// TIA Portal project "batch Steam cooker V2" (V19)

(* hardware
DEVICE "S7-1200 station_1"  S7-1200 Station
   slot 0: "Rack_0"  S7-1200 Rack  Rack  V1.0
   slot 1: "PLC_1"  CPU 1214C AC/DC/Rly  6ES7 214-1BG40-0XB0  V4.5
DEVICE "HMI_2"  TP700 Comfort
   slot 0: "HMI_2"  TP700 Comfort  6AV2 124-0GC01-0AX0  17.0.0.0
   slot 1: "HMI_RT_2"  TP700 Comfort  6AV2 124-0GC01-0AX0  17.0.0.0
   slot 5: "HMI_2.IE_CP_1"  PROFINET Interface  17.0.0.0
      slot 1: "PROFINET Interface_1"  PROFINET Interface
         slot 1: "Port_1"  Port
         slot 2: "Port_2"  Port
   slot 7: "HMI_2.MPI/DP_CP_1"  MPI/DP Interface  17.0.0.0
*)

// ===== PLC "PLC_1"  CPU 1214C AC/DC/Rly =====

VAR_GLOBAL   // PLC tag table "Default tag table"
   "Vacuum Pump Starter" AT %Q4.0 : Bool;
   "Steam Regulator" AT %Q4.1 : Bool;
   "Cooling Water Valve" AT %Q4.2 : Bool;
   "Green Light" AT %Q3.0 : Bool;
   "Red Light" AT %Q3.2 : Bool;
   "Yellow Light" AT %Q3.1 : Bool;
   "Alarm_Word" AT %MW3 : Int;
   "Tag_1" AT %M3.0 : Bool;
   "Tag_2" AT %M3.1 : Bool;
   "Tag_3" AT %M3.6 : Bool;
   "Tag_4" AT %M3.7 : Bool;
   "Tag_5" AT %M4.0 : Bool;
   "Tag_6" AT %M4.1 : Bool;
   "Tag_7" AT %M3.2 : Bool;
   "Tag_8" AT %M3.3 : Bool;
   "Tag_9" AT %M3.4 : Bool;
   "Tag_10" AT %M3.5 : Bool;
   "Acknowledge_Word" AT %MW4 : Int;
   "Acknowledge bit" AT %M5.0 : Bool;
END_VAR

VAR_GLOBAL   // PLC tag table "IO_Inputs"
   "Door Lock FB" AT %I0.1 : Bool;
   "Manhole Closed FB" AT %I0.2 : Bool;
   "Manhole Open FB" AT %I0.3 : Bool;
   "Water Level FB" AT %I0.4 : Bool;
   "Door Interlock" AT %I0.5 : Bool;
   "Emergency Stop" AT %I0.7 : Bool;
   "Pressure Input" AT %ID68 : Real;
   "Temperature Input" AT %ID64 : Real;
   "Water Flow Input" AT %ID72 : Real;
END_VAR

VAR_GLOBAL   // PLC tag table "IO_Outputs"
   "V1 Output" AT %Q0.0 : Bool;
   "V2 Output" AT %Q0.1 : Bool;
   "V3 Output" AT %Q0.2 : Bool;
   "V9" AT %Q1.0 : Bool;
   "V8" AT %Q0.7 : Bool;
   "V7" AT %Q0.6 : Bool;
   "V6" AT %Q0.5 : Bool;
   "V5" AT %Q0.4 : Bool;
   "V4" AT %Q0.3 : Bool;
   "Motor Run Output" AT %Q2.0 : Bool;
   "Motor Direction Output" AT %Q2.1 : Bool;
END_VAR

VAR_GLOBAL CONSTANT   // PLC tag table "Const"
   "cIdle" : Int := 50;
   "cLock" : Int := 15;
   "cAddWater" : Int := 1;
   "cOpenMH" : Int := 2;
   "cWaitMat" : Int := 3;
   "cCloseMH" : Int := 4;
   "cColdMix" : Int := 5;
   "cHeat" : Int := 6;
   "cCook" : Int := 7;
   "cConfDis" : Int := 10;
   "cDisch" : Int := 11;
   "cFinal" : Int := 12;
END_VAR

TYPE "UDT_Recipe_Production"
   STRUCT
      Recipe_Name : String := 'DEFAULT';   // Recipe identification name
      Recipe_Number : UInt := 1;   // Recipe ID number (1-99)
      Heating_Temp_Phase1 : Real := 80.0;   // Cooking temperature setpoint (°C)
      Adding_Water1_QTY : Real := 100.0;   // First water addition quantity (Liters)
      Cold_Mix_Time : Time := T#300S;   // Cold mix time before heating (seconds)
      Cooking_Time_Phase1 : Time := T#1800S;   // Cooking time after temp reached (seconds)
      Compensation_Time : Time := T#600S;   // Additional processing time (seconds)
      Discharge_Time : Time;   // Auto discharge time (0=manual only)
      Water_Flow_Timeout : Time := T#120S;   // Water addition timeout
      Manhole_Open_Time : Time :=  T#30S;   // Manhole opening timeout
      Manhole_Close_Time : Time :=  T#30S;   // Manhole closing timeout
      Steam_Ramp_Rate : Real := 5.0;   // Steam valve opening rate %/sec
      Vacuum_Enable : Bool := true;   // Enable vacuum during cooking
      Final_Temp_Target : Real := 75.0;   // Final product temperature (°C)
      Product_Type : UInt := 1;   // Product type (1=Soft, 2=Hard, 3=Special)
      Batch_Size_kg : Real := 300.0;
   END_STRUCT;
END_TYPE

TYPE "UDT_Motor_Command"
   STRUCT
      Priority : UInt := 0;   // Command priority (1=Auto, 2=Func, 3=Man)
      Start_Man : Bool;
      Start_Func : Bool;
      Start_Auto : Bool;
      Stop : Bool;
      Reset : Bool;
      Pulse_Enable : Bool;
      Discharge_Mode : Bool;
      Enable : Bool;
      Direction : Int;
      Speed_SP_pct : Real;   // Speed setpoint %
   END_STRUCT;
END_TYPE

TYPE "UDT_Motor_Config"
   STRUCT
      Motor_Name : String;
      Max_Speed_pct : Real := 100.0;
      Min_Speed_pct : Real := 0.0;
      Start_Timeout : Time := T#10S;
      Stop_Timeout : Time := T#5S ;
      Rev_Dwell : Time := T#2S ;   // Direction change dwell
      T_Fwd : Time := T#30S ;
      T_Hold : Time := T#5S ;
      T_Bwd : Time := T#20S ;
      Disch_Speed_pct : Real := 25.0;
      Acceleration_Time : Time := T#3S;
      Deceleration_Time : Time := T#3S;
      Interlock_Used : Bool := TRUE;
      Motor_Type : UInt := 1;
      Rated_Speed_RPM : Real;
      Rated_Power_kW : Real;
   END_STRUCT;
END_TYPE

TYPE "UDT_Motor_Status"
   STRUCT
      Running : Bool;   // Motor is running
      Fault : Bool;
      Fault_Code : UInt;
      Direction : UInt;   // Direction (0=Stop, 1=Fwd, 2=Rev)
      State : UInt;   // State (0=Stop, 1=Fwd, 2=Hold, 3=Bwd)
      Source : UInt;   // Command source (0=None, 1=Auto, 2=Func, 3=Man)
      Ready : Bool;
      Position_pct : Real;   // Position feedback %
      Speed_Actual_pct : Real;
      Runtime_Hours : Real;
      Start_Count : UDInt;
      R_Fwd : Bool;
      R_Rev : Bool;
      RDwell_Q : Bool;
   END_STRUCT;
END_TYPE

TYPE "UDT_Motor_Outputs"
   STRUCT
      Q_Run : Bool;
      Q_DirFwd : Bool;
      Q_Stop : Bool;
      Contactor_Main : Bool;
      Contactor_Star : Bool;
      Contactor_Delta : Bool;
      Brake_Release : Bool;
      Alarm_Output : Bool;
      Status_LED : UInt;
      AO_SpeedPct : Real;
      AO_Torque : Real;
   END_STRUCT;
END_TYPE

TYPE "UDT_Motor_Interlocks"
   STRUCT
      Permissive : Bool := true;   // General permissive
      OOS : Bool;   // Out of service
      E_Stop : Bool;
      Drive_Ready : Bool;   // Drive ready feedback
      Drive_Fault : Bool;
      Temperature_OK : Bool := true;
      Vibration_OK : Bool := true;
      Overcurrent_OK : Bool := true;
      Door_Closed : Bool := TRUE;
      Guard_OK : Bool := TRUE;
      Lubrication_OK : Bool := TRUE;
      Cooling_OK : Bool := TRUE;
      Local_Stop : Bool;
      Drive_Running : Bool;
      Overload : Bool;
      VFD_Fault : Bool;
   END_STRUCT;
END_TYPE

TYPE "UDT_Motor"
   STRUCT
      Command : "UDT_Motor_Command";
      Outputs : "UDT_Motor_Outputs";   // Physical outputs
      Config : "UDT_Motor_Config";
      Status : "UDT_Motor_Status";
      Interlocks : "UDT_Motor_Interlocks";
   END_STRUCT;
END_TYPE

TYPE "UDT_Valve_Command"
   STRUCT
      Priority : UInt;
      Open_Man : Bool;
      Open_Auto : Bool;
      Close_Auto : Bool;
      Close_Man : Bool;
      Open_Func : Bool;
      Close_Func : Bool;
      Reset : Bool;
      Emergency_Close : Bool;
   END_STRUCT;
END_TYPE

TYPE "UDT_Valve_Config"
   STRUCT
      Valve_Type : UInt := 1;
      Valve_Name : String;
      Travel_Timeout : Time := T#30ms;
      Stroke_Time : Time := T#15ms;
      Position_Tolerance : Real := 2.0;
      Min_Position : Real;
      Max_Position : Real := 100.0;
      Fail_Position : UInt;
      TwoCoils : Bool;
      Actuator_Type : UInt := 1;
      Feedback_Type : UInt := 1;
      Service_Hours : Real;
      Interlock_Used : Bool := True;
      Fail_Safe_Position : Bool;
      Open_Time : Time;
      Close_Time : Time;
   END_STRUCT;
END_TYPE

TYPE "UDT_Valve_Status"
   STRUCT
      Fault : Bool;
      Fault_Code : UInt;
      State : UInt;   // State (0=Stop, 1=Fwd, 2=Hold, 3=Bwd)
      Source : UInt;   // Command source (0=None, 1=Auto, 2=Func, 3=Man)
      Ready : Bool;
      Moving : Bool;
      At_Position : Bool;
      Travel_Time : Time;
      Operation_Count : UDInt;
      Position_Actual_pct : Real;   // Position feedback %
      Runtime_Hours : Real;
      Limit_Open : Bool;
      Limit_Closed : Bool;
      Open : Bool;
      Closed : Bool;
   END_STRUCT;
END_TYPE

TYPE "UDT_Valve_Outputs"
   STRUCT
      Q_Run : Bool;
      Q_Open : Bool;
      Q_Close : Bool;
      Solenoid_A : Bool;
      Solenoid_B : Bool;
      Motor_CW : Bool;
      Motor_CCW : Bool;
      Brake_Release : Bool;
      Status_LED : Bool;
      Alarm_Output : Bool;
      AO_Position_pct : Real;
   END_STRUCT;
END_TYPE

TYPE "UDT_Valve_Interlocks"
   STRUCT
      Permissive : Bool := true;   // General permissive
      OOS : Bool;   // Out of service
      E_Stop : Bool;
      Process_Temp_OK : Bool := true;
      Local_Isolation : Bool;
      Process_Pressure_OK : Bool := TRUE        ;
      Upstream_OK : Bool := TRUE        ;
      Downstream_OK : Bool := TRUE        ;
      Interlock_Chain : Bool := TRUE        ;
      Maintenance_Lock : Bool;
      Air_Pressure_OK : Bool := TRUE        ;
      Power_Available : Bool := TRUE        ;
   END_STRUCT;
END_TYPE

TYPE "UDT_Valve"
   STRUCT
      Command : "UDT_Valve_Command";
      Config : "UDT_Valve_Config";
      Status : "UDT_Valve_Status";
      Outputs : "UDT_Valve_Outputs";
      Interlocks : "UDT_Valve_Interlocks";
      Open_Auto : Bool;
      Priority : UInt;
      Reset : Bool;
      Open_Man : Bool;
      Close_Man : Bool;
      Open_Func : Bool;
      Close_Func : Bool;
      Close_Auto : Bool;
      Position_SP_pct : Real;
      Enable : Bool;
      Emergency_Close : Bool;
   END_STRUCT;
END_TYPE

TYPE "UDT_Recipe_Screw"
   STRUCT
      Forward_Speed_pct : Real := 75.0;   // Forward screw speed %
      Backward_Speed_pct : Real := 50.0;
      Reverse_Speed_pct : Real := 50.0;
      Forward_Run_Time : Time := T#30S ;   // Forward running time (pulsing)
      Backward_Run_Time : Time := T#20S ;
      Hold_Time : Time := T#10S ;   // Hold time between direction changes
      Pause_Time : Time := T#5S ;   // Pause between pulse cycles
      Direction_Change_Delay : Time := T#2S;   // Delay between direction changes
      Screw_Ramp_Time : Time := T#3S;   // Speed ramp up/down time
      Max_Runtime_Continuous : Time := T#600S;   // Max continuous runtime before pause
      Discharge_Speed_pct : Real := 25.0;   // Screw speed during discharge %
      Cold_Mix_Speed_pct : Real := 60.0;   // Speed during cold mixing %
      Cook_Mix_Speed_pct : Real := 80.0;   // Speed during cooking phase %
      Pulse_Enable_ColdMix : Bool := TRUE;   // Enable pulsing during cold mix
      Pulse_Enable_Cooking : Bool := TRUE;
      Pulse_Enable_Discharge : Bool;
      Pulse_Time_On : Time;
      Pulse_Time_Off : Time;
   END_STRUCT;
END_TYPE

TYPE "UDT_Recipe_Temperature"
   STRUCT
      Heat_Setpoint_Phase1 : Real := 80.0;
      Heat_Setpoint_Phase2 : Real := 85.0;
      Heat_Deadband : Real := 2.0;
      Heat_Rate_Limit : Real := 2.0;
      Cool_Setpoint : Real := 60.0;
      Cool_Rate_Limit : Real := 1.0;
      Steam_Pressure_Max : Real := 6.0;
      Steam_Pressure_Min : Real := 2.0;
      Temp_Alarm_High : Real := 95.0;
      Temp_Alarm_Low : Real := 40.0;
      Temp_Sensor_Timeout : Time := T#10S;
      Heat_Timeout : Time := T#1800S;
      Cool_Timeout : Time := T#900S;
      Overtemp_Shutdown : Real := 100.0;
      Cool_Deadband : Real;
   END_STRUCT;
END_TYPE

TYPE "UDT_Recipe_Vacuum"
   STRUCT
      Vacuum_Setpoint_mbar : Real := 500.0;   // Vacuum setpoint (mbar absolute)
      Vacuum_Tolerance : Real := 50.0;   // Vacuum tolerance (±mbar)
      Vacuum_Offset_pct : Real := 5.0;   // Hysteresis offset percentage
      Pump_Start_Delay : Time := T#5S;   // Pump start delay after valve open
      Pump_Stop_Delay : Time := T#10S;   // Pump stop delay after valve close
      Max_Vacuum_Time : Time := T#3600S;   // aximum continuous vacuum time
      Vacuum_Break_Pressure : Real := 900.0;   // Vacuum break pressure (mbar)
      Leak_Test_Time : Time := T#60S;   // Vacuum leak test duration
      Leak_Test_Tolerance : Real := 10.0;   // Acceptable leak rate (mbar/min)
      Emergency_Break_Enable : Bool := TRUE;   // Enable emergency vacuum break
      Cooling_Vacuum_Enable : Bool := TRUE;   // Enable vacuum during cooling
      Cooking_Vacuum_Enable : Bool;
      Vacuum_Pump_Timeout : Time := T#30S;   // Vacuum pump start timeout
      Pressure_Sensor_Timeout : Time := T#10S;   // Pressure sensor timeout
      Min_Vacuum_Quality : Real := 100.0;   // Minimum vacuum level (mbar)
   END_STRUCT;
END_TYPE

TYPE "UDT_Recipe_Complete"
   STRUCT
      Production : "UDT_Recipe_Production";   // Production parameters
      Screw : "UDT_Recipe_Screw";
      Temperature : "UDT_Recipe_Temperature";
      Vacuum : "UDT_Recipe_Vacuum";
      Recipe_Valid : Bool;
      Recipe_Locked : Bool;
      Creation_Date : DTL;
      Modified_Date : DTL;
      Created_By : String := 'SYSTEM';
      Modified_By : String := 'SYSTEM';
      Recipe_Version : Real := 1.0;
      Recipe_Notes : String;
   END_STRUCT;
END_TYPE

TYPE "UDT_Process_Status"
   STRUCT
      Current_Step : UInt := 50;
      Step_Name : String := 'IDLE';
      Phase_Name : String := 'IDLE';
      Phase_Active : UInt;   // Active phase (0=Idle, 1=Prep, 2=Mix, 3=Cook, 4=Discharge)
      Current_Phase : UInt;
      Time_Remaining : Time;
      Time_Elapsed : Time;
      Total_Batch_Time : Time;
      Step_Progress_pct : Real;
      Batch_Progress_pct : Real;
      Temp_Actual : Real := 25.0;
      Temp_Setpoint : Real;
      Pressure_Actual : Real := 1013.0;
      Pressure_Setpoint : Real;   // Current pressure setpoint (mbar)
      Water_Level_Actual : Real;
      Water_Level_Target : Real;
      Screw_Speed_Actual : Real;
      Screw_Speed_Setpoint : Real;   // Screw speed setpoint %
      Batch_Number : UInt := 1;   // Current water level (L)
      Recipe_Active : UInt := 1;
      Process_Running : Bool;
      Process_Paused : Bool;
      Process_Complete : Bool;
      Process_Aborted : Bool;
      Fault_Active : Bool;   // System fault active flag
      Emergency_Stop : Bool;   // Emergency stop active flag
      Operator_Present : Bool;   // Operator attention required
      System_Ready : Bool;
      Overall_Progress : Real;
      Individual_Discharge_Active : Bool;
   END_STRUCT;
END_TYPE

TYPE "UDT_Process_HMI"
   STRUCT
      Start_Production : Bool;
      Stop_Production : Bool;
      Reset_System : Bool;
      Reset_p_s : Bool;
      Abort_Process : Bool;
      Acknowledge_Alarms : Bool;
      RawMaterial_OK : Bool;
      Manhole_Secured_OK : Bool;
      Discharge_Ready_OK : Bool;
      Quality_Check_OK : Bool;
      Cleaning_Complete_OK : Bool;
      Recipe_Selected : UInt := 1;
      Load_Recipe : Bool;
      Save_Recipe : Bool;
      Recipe_Edit_Mode : Bool;
      Recipe_Backup : Bool;
      Recipe_Restore : Bool;
      Manual_ON : Array[0..15] of Bool;   // Manual ON commands [V1-V9, R1, Aux1-5]
      Manual_OFF : Array[0..15] of Bool;
      Auto_Mode : Array[0..15] of Bool;
      Temp_Override_Enable : Bool;
      Temp_Override_Value : Real;
      Speed_Override_Enable : Bool;
      Speed_Override_Value : Real;
      Time_Override_Enable : Bool;
      Time_Override_Factor : Real := 1.0;
      Operator_ID : String := 'UNKNOWN';
      Shift_ID : UInt := 1;
      Production_Mode : UInt := 1;   // Mode (1=Auto, 2=Manual, 3=Test)
      System_Ready : Bool;
      Maintenance_Mode : Bool;
      Individual_Discharge_Button : Bool;
   END_STRUCT;
END_TYPE

TYPE "UDT_Process_IO"
   STRUCT
      FS_Water_Flow : Bool;
      LS1_Discharge_Locked : Bool;
      LS2_Manhole_Closed : Bool;
      LS3_Manhole_Opened : Bool;
      LL_Water_Level : Bool;
      ES_Emergency_Stop : Bool;
      PS_Steam_Pressure_OK : Bool;
      PS_Air_Pressure_OK : Bool;
      TS_Steam_Temperature_OK : Bool;
      Door_Interlock_OK : Bool;
      Guard_Switch_OK : Bool;
      Door_Locked_FB : Bool;
      Door_Unlocked_FB : Bool;
      Water_Level_FB : Bool;
      Manhole_Open_FB : Bool;
      Manhole_Closed_FB : Bool;
      AI_Temperature : Real := 25.0;
      AI_Pressure : Real := 1013.0;
      AI_Steam_Pressure : Real;
      AI_Water_Flow : Real;
      AI_Steam_Flow : Real;
      AI_Vacuum_Level : Real := 1013.0;
      AI_Motor_Current : Real;
      AI_Motor_Power : Real;
      DO_Alarm_Horn : Bool;
      DO_Status_Green : Bool;
      DO_Status_Yellow : Bool;
      DO_Status_Red : Bool;
      DO_Vacuum_Pump : Bool;   // Vacuum pump starter (K1)
      DO_Steam_Regulator_En : Bool;
      DO_Cooling_Water : Bool;
      DO_Process_Light : Bool;
      AO_Steam_Regulator : Real;
      AO_Cooling_Control : Real;
      AO_Process_Speed : Real;
   END_STRUCT;
END_TYPE

DATA_BLOCK "DB_Recipes"   // DB1
{ S7_Optimized_Access := 'TRUE' }
VERSION : 0.1
   VAR
      Recipes : Array[1..10] of "UDT_Recipe_Complete";   // Recipe storage array (1-10)
      Active_Recipe : "UDT_Recipe_Complete";   // Currently loaded recipe
      Default_Recipe : "UDT_Recipe_Complete";   // Factory default recipe
   END_VAR
BEGIN
   Default_Recipe.Production.Recipe_Name := 'DEFAULT_CHEESE';
   Default_Recipe.Production.Batch_Size_kg := 1000.0;
   Default_Recipe.Production.Adding_Water1_QTY := 100.0;
   Default_Recipe.Production.Water_Flow_Timeout := T#120S;
   Default_Recipe.Production.Cold_Mix_Time := T#300S;
   Default_Recipe.Production.Cooking_Time_Phase1 := T#1800S;
   Default_Recipe.Production.Heating_Temp_Phase1 := 80.0;
   Default_Recipe.Screw.Cold_Mix_Speed_pct := 60.0;
   Default_Recipe.Screw.Cook_Mix_Speed_pct := 80.0;
   Default_Recipe.Screw.Discharge_Speed_pct := 25.0;
   Default_Recipe.Temperature.Heat_Setpoint_Phase1 := 80.0;
   Default_Recipe.Temperature.Heat_Deadband := 2.0;
   Default_Recipe.Temperature.Heat_Timeout := T#1800S;
   Default_Recipe.Recipe_Valid := TRUE;
   Default_Recipe.Production.Recipe_Number := 1;
   Default_Recipe.Production.Manhole_Open_Time := T#30S;
   Default_Recipe.Production.Manhole_Close_Time := T#30S;
   Default_Recipe.Screw.Pulse_Enable_ColdMix := TRUE;
   Default_Recipe.Screw.Pulse_Enable_Cooking := TRUE;
   Default_Recipe.Vacuum.Vacuum_Setpoint_mbar := 500.0;
   Default_Recipe.Vacuum.Vacuum_Tolerance := 50.0;
   Default_Recipe.Vacuum.Cooking_Vacuum_Enable := FALSE;
   Active_Recipe.Production.Water_Flow_Timeout := T#10S;
   Active_Recipe.Production.Compensation_Time := T#6S;
   Active_Recipe.Production.Cooking_Time_Phase1 := T#10S;
   Active_Recipe.Production.Cold_Mix_Time := T#20S;
   Active_Recipe.Production.Discharge_Time := T#6ms;
   Active_Recipe.Vacuum.Cooking_Vacuum_Enable := TRUE;
END_DATA_BLOCK

DATA_BLOCK "FB_Process_Main_DB"   // DB2
{ S7_Optimized_Access := 'TRUE' }
VERSION : 0.1
// stored: InstanceOfName FB_Process_Main
"FB_Process_Main"
BEGIN
END_DATA_BLOCK

DATA_BLOCK "FB_Motor_VFD_DB_1"   // DB3
{ S7_Optimized_Access := 'TRUE' }
VERSION : 0.1
// stored: InstanceOfName FB_Motor_VFD
"FB_Motor_VFD"
BEGIN
END_DATA_BLOCK

DATA_BLOCK "FB_Motor_VFD_DB"   // DB13
{ S7_Optimized_Access := 'TRUE' }
VERSION : 0.1
// stored: InstanceOfName FB_Motor_VFD
"FB_Motor_VFD"
BEGIN
END_DATA_BLOCK

DATA_BLOCK "ALarms"   // DB14
{ S7_Optimized_Access := 'TRUE' }
VERSION : 0.1
   VAR
      Alarms : UInt;
   END_VAR
BEGIN
END_DATA_BLOCK

DATA_BLOCK "FB_Valve_DO_DB"   // DB15
{ S7_Optimized_Access := 'TRUE' }
VERSION : 0.1
// stored: InstanceOfName FB_Valve_DO
"FB_Valve_DO"
BEGIN
END_DATA_BLOCK

DATA_BLOCK "DB_Motors"   // DB18
{ S7_Optimized_Access := 'TRUE' }
VERSION : 0.1
   VAR RETAIN
      Motors : Array[1..1] of "UDT_Motor";   // Motor control array - =Screw Motor
   END_VAR
BEGIN
   Motors[1].Config.Motor_Name := 'SCREW_MOTOR';
   Motors[1].Config.Max_Speed_pct := 1800.0;
   Motors[1].Config.Rated_Speed_RPM := 1800.0;
   Motors[1].Config.Rated_Power_kW := 15.0;
   Motors[1].Config.Acceleration_Time := T#10S;
   Motors[1].Config.Rev_Dwell := T#2S;
   Motors[1].Config.Disch_Speed_pct := 25.0;
   Motors[1].Config.Start_Timeout := T#10S;
   Motors[1].Config.T_Fwd := T#30S;
   Motors[1].Config.T_Hold := T#5S;
   Motors[1].Config.T_Bwd := T#20S;
END_DATA_BLOCK

DATA_BLOCK "DB_Valves"   // DB19
{ S7_Optimized_Access := 'TRUE' }
VERSION : 0.1
   VAR
      Valves : Array[1..9] of "UDT_Valve";   // Valve control array - =V1 Manhole, =V2 CIP, ..., =V9 Vacuum Cooling
   END_VAR
BEGIN
   Valves[1].Config.Valve_Name := 'V1_MANHOLE';
   Valves[2].Config.Valve_Name := 'V2_CIP';
   Valves[3].Config.Valve_Name := 'V3_DISCHARGE_UNLOCK';
   Valves[4].Config.Valve_Name := 'V4_DISCHARGE';
   Valves[5].Config.Valve_Name := 'V5_WATER';
   Valves[6].Config.Valve_Name := 'V6_STEAM';
   Valves[7].Config.Valve_Name := 'V7_EVACUATION';
   Valves[8].Config.Valve_Name := 'V8_VACUUM';
   Valves[9].Config.Valve_Name := 'V9_VACUUM_COOLING';
   Valves[1].Config.Travel_Timeout := T#30S;
   Valves[2].Config.Travel_Timeout := T#15S;
   Valves[3].Config.Travel_Timeout := T#30S;
   Valves[4].Config.Travel_Timeout := T#20S;
   Valves[5].Config.Travel_Timeout := T#15S;
   Valves[6].Config.Travel_Timeout := T#10S;
   Valves[7].Config.Travel_Timeout := T#15S;
   Valves[8].Config.Travel_Timeout := T#20S;
   Valves[9].Config.Travel_Timeout := T#15S;
END_DATA_BLOCK

DATA_BLOCK "DB_Test_Motors"   // DB20
{ S7_Optimized_Access := 'FALSE' }
VERSION : 0.1
   VAR
      ff : Int;
   END_VAR
BEGIN
END_DATA_BLOCK

DATA_BLOCK "DB_Process"   // DB21
{ S7_Optimized_Access := 'FALSE' }
VERSION : 0.1
   VAR
      Status : "UDT_Process_Status";   // current process
      HMI : "UDT_Process_HMI";
      IO : "UDT_Process_IO";
      Timers : Array[1..10] of TON_TIME;
      Counters : Array[1..5] of CTU_INT;
   END_VAR
BEGIN
   Status.Current_Step := 50;
   Status.Step_Name := 'IDLE';
   Status.Batch_Number := 1;
   Status.Recipe_Active := 1;
   HMI.Shift_ID := 1;
   HMI.Operator_ID := 'OPERATOR';
   IO.AI_Pressure := 1000.0;
   IO.AI_Steam_Pressure := 25.0;
   IO.Manhole_Open_FB := true;
END_DATA_BLOCK

FUNCTION_BLOCK "FB_Valve_DO"   // FB1, LAD
{ S7_Optimized_Access := 'TRUE' }
VERSION : 0.1
   VAR_INPUT
      AutoCmd : Bool;   // from automatic sequence (open=TRUE)
      FuncCmd : Bool;   // from Function screens
      ManCmd : Bool;   // from Manual page (your ON/OFF button drives this)
      OOS : Bool;   // Out Of Service; forces closed
      Permissive : Bool;   // E‑Stop OK, interlocks OK
      FbOpen : Bool;   // optional open limit switch
      FbClosed : Bool;   // optional closed limit switch
      TwoCoils : Bool;   // TRUE = separate open/close coils; FALSE = single coil
      T_Stroke : Time := T#3S;   // normal movement time (e.g., T#5S)
      T_Timeout : Time := T#6S;   // fault timeout (e.g., T#10S)
   END_VAR
   VAR_OUTPUT
      Q_Open : Bool;   // open (or single) coil
      Q_Close : Bool;   // close coil (only used if TwoCoils=TRUE)
      Ready : Bool;
      FaultTO : Bool;
      FaultFB : Bool;
      Source : UInt;   // 1 Auto, 2 Func, 3 Man
      Status : UInt;   // 0 Unknown, 1 Closed, 2 Opening, 3 Open, 4 Closing, 5 Fault
   END_VAR
   VAR
      Cmd_DesiredOpen_raw : Bool;
      Cmd_DesiredOpen_OK : Bool;
      Req_Open : Bool;
      Req_Close : Bool;
      St_Opening : Bool;
      St_Closing : Bool;
      St_Open : Bool;
      St_Closed : Bool;
      St_Moving : Bool;
      Open_Reached : Bool;
      Close_Reached : Bool;
      FaultLatched : Bool;
      TON_Move : TON_TIME;
      TON_Timeout : TON_TIME;
   END_VAR
   VAR_TEMP
      MoveEnable : Bool;
   END_VAR
BEGIN

REGION Network 1: Conflict for feedback
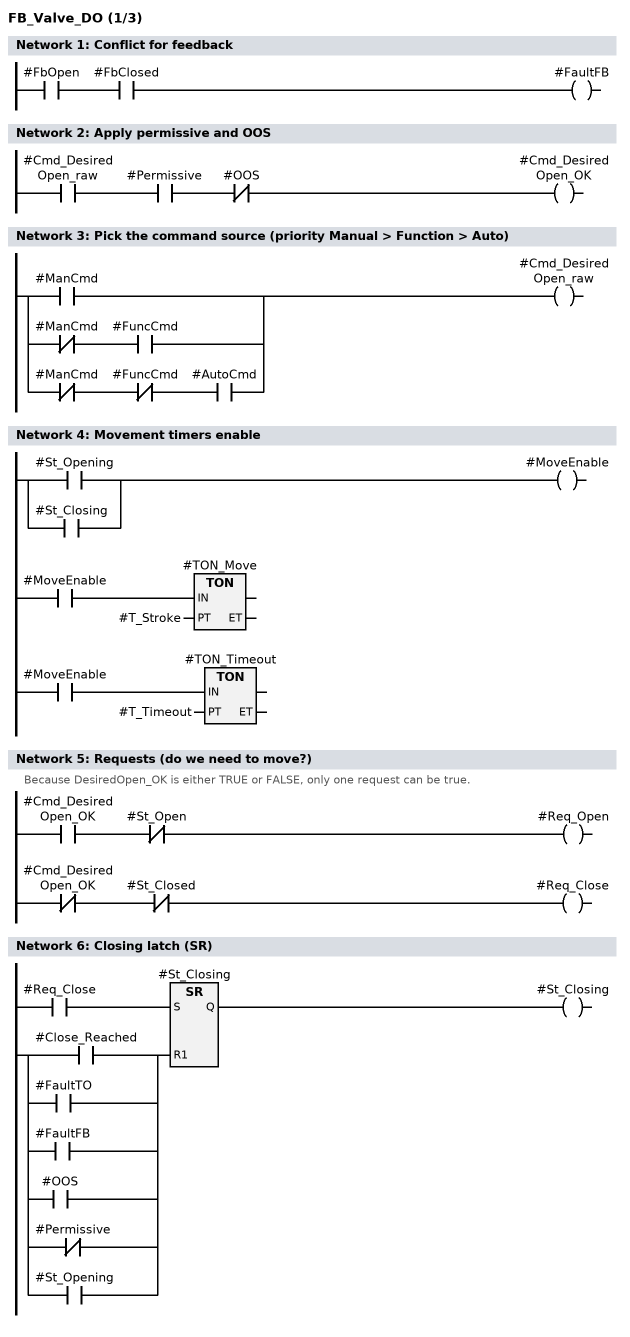
   RUNG wire#powerrail
      Contact( #FbOpen )
      Contact( #FbClosed )
      Coil( #FaultFB )
   END_RUNG
   // the same network as SCL:
   #FaultFB := #FbOpen AND #FbClosed;
END_REGION

REGION Network 2: Apply permissive and OOS
   RUNG wire#powerrail
      Contact( #Cmd_DesiredOpen_raw )
      Contact( #Permissive )
      I_Contact( #OOS )
      Coil( #Cmd_DesiredOpen_OK )
   END_RUNG
   // the same network as SCL:
   #Cmd_DesiredOpen_OK := #Cmd_DesiredOpen_raw AND #Permissive AND NOT #OOS;
END_REGION

REGION Network 3: Pick the command source (priority Manual > Function > Auto)
   RUNG wire#powerrail
      Contact( #ManCmd )
      wire#w1
      Coil( #Cmd_DesiredOpen_raw )
   END_RUNG
   RUNG wire#powerrail
      I_Contact( #ManCmd )
      Contact( #FuncCmd )
   END_RUNG wire#w1
   RUNG wire#powerrail
      I_Contact( #ManCmd )
      I_Contact( #FuncCmd )
      Contact( #AutoCmd )
   END_RUNG wire#w1
   // the same network as SCL:
   #Cmd_DesiredOpen_raw := #ManCmd OR (NOT #ManCmd AND #FuncCmd) OR (NOT #ManCmd AND NOT #FuncCmd AND #AutoCmd);
END_REGION

REGION Network 4: Movement timers enable
   #MoveEnable := #St_Opening OR #St_Closing;
   #TON_Move(IN := #MoveEnable, PT := #T_Stroke);   // TON
   #TON_Timeout(IN := #MoveEnable, PT := #T_Timeout);   // TON
END_REGION

REGION Network 5: Requests (do we need to move?)
   // Because DesiredOpen_OK is either TRUE or FALSE, only one request can be true.
   RUNG wire#powerrail
      Contact( #Cmd_DesiredOpen_OK )
      I_Contact( #St_Open )
      Coil( #Req_Open )
   END_RUNG
   RUNG wire#powerrail
      I_Contact( #Cmd_DesiredOpen_OK )
      I_Contact( #St_Closed )
      Coil( #Req_Close )
   END_RUNG
   // the same network as SCL:
   #Req_Open := #Cmd_DesiredOpen_OK AND NOT #St_Open;
   #Req_Close := NOT #Cmd_DesiredOpen_OK AND NOT #St_Closed;
END_REGION

REGION Network 6: Closing latch (SR)
   RUNG wire#powerrail
      Contact( #Req_Close )
      S_SR(operand := #St_Closing, r1 := wire#w1)
      Coil( #St_Closing )
   END_RUNG
   RUNG wire#powerrail
      Contact( #Close_Reached )
   END_RUNG wire#w1
   RUNG wire#powerrail
      Contact( #FaultTO )
   END_RUNG wire#w1
   RUNG wire#powerrail
      Contact( #FaultFB )
   END_RUNG wire#w1
   RUNG wire#powerrail
      Contact( #OOS )
   END_RUNG wire#w1
   RUNG wire#powerrail
      I_Contact( #Permissive )
   END_RUNG wire#w1
   RUNG wire#powerrail
      Contact( #St_Opening )
   END_RUNG wire#w1
   // the same network as SCL:
   IF #Req_Close THEN
       #St_Closing := TRUE;   // SR flip-flop
   END_IF;
   IF #Close_Reached OR #FaultTO OR #FaultFB OR #OOS OR NOT #Permissive OR #St_Opening THEN
       #St_Closing := FALSE;
   END_IF;
   #St_Closing := #St_Closing;
END_REGION

REGION Network 7: Latch “Opening” (SR)
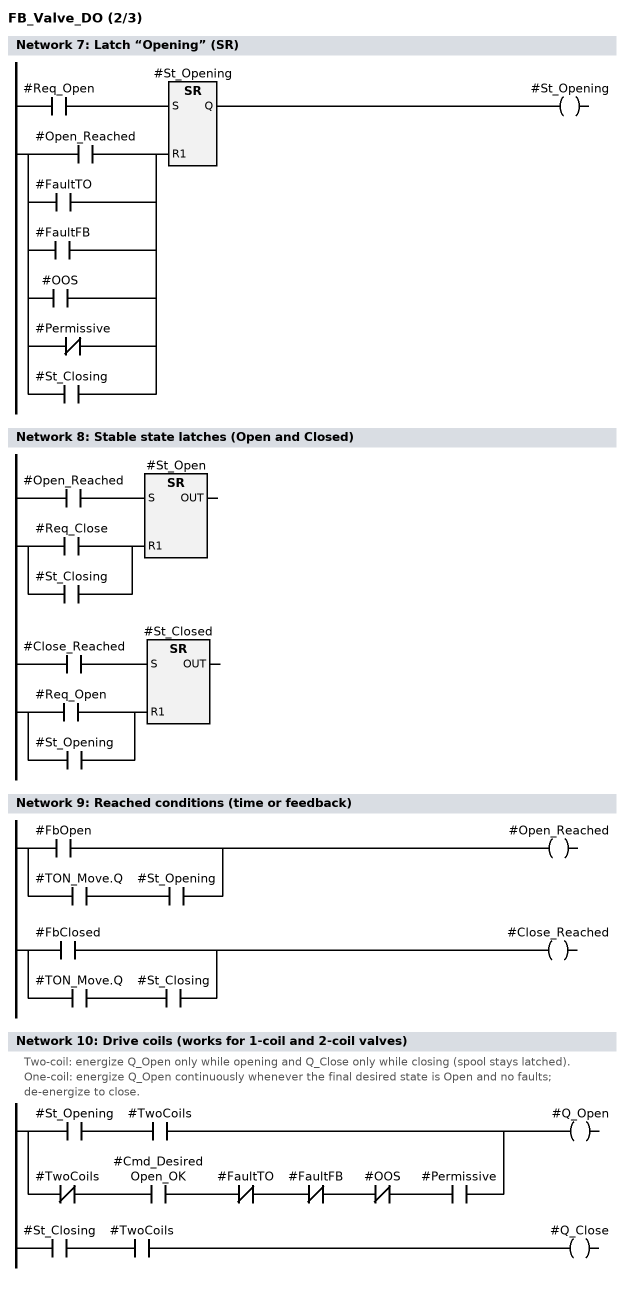
   RUNG wire#powerrail
      Contact( #Req_Open )
      S_SR(operand := #St_Opening, r1 := wire#w1)
      Coil( #St_Opening )
   END_RUNG
   RUNG wire#powerrail
      Contact( #Open_Reached )
   END_RUNG wire#w1
   RUNG wire#powerrail
      Contact( #FaultTO )
   END_RUNG wire#w1
   RUNG wire#powerrail
      Contact( #FaultFB )
   END_RUNG wire#w1
   RUNG wire#powerrail
      Contact( #OOS )
   END_RUNG wire#w1
   RUNG wire#powerrail
      I_Contact( #Permissive )
   END_RUNG wire#w1
   RUNG wire#powerrail
      Contact( #St_Closing )
   END_RUNG wire#w1
   // the same network as SCL:
   IF #Req_Open THEN
       #St_Opening := TRUE;   // SR flip-flop
   END_IF;
   IF #Open_Reached OR #FaultTO OR #FaultFB OR #OOS OR NOT #Permissive OR #St_Closing THEN
       #St_Opening := FALSE;
   END_IF;
   #St_Opening := #St_Opening;
END_REGION

REGION Network 8: Stable state latches (Open and Closed)
   RUNG wire#powerrail
      Contact( #Open_Reached )
      S_SR(operand := #St_Open, r1 := wire#w1)
   END_RUNG
   RUNG wire#powerrail
      Contact( #Req_Close )
   END_RUNG wire#w1
   RUNG wire#powerrail
      Contact( #St_Closing )
   END_RUNG wire#w1
   RUNG wire#powerrail
      Contact( #Close_Reached )
      S_SR(operand := #St_Closed, r1 := wire#w2)
   END_RUNG
   RUNG wire#powerrail
      Contact( #Req_Open )
   END_RUNG wire#w2
   RUNG wire#powerrail
      Contact( #St_Opening )
   END_RUNG wire#w2
   // the same network as SCL:
   IF #Open_Reached THEN
       #St_Open := TRUE;   // SR flip-flop
   END_IF;
   IF #Req_Close OR #St_Closing THEN #St_Open := FALSE; END_IF;
   IF #Close_Reached THEN
       #St_Closed := TRUE;   // SR flip-flop
   END_IF;
   IF #Req_Open OR #St_Opening THEN #St_Closed := FALSE; END_IF;
END_REGION

REGION Network 9: Reached conditions (time or feedback)
   RUNG wire#powerrail
      Contact( #FbOpen )
      wire#w1
      Coil( #Open_Reached )
   END_RUNG
   RUNG wire#powerrail
      Contact( #TON_Move.Q )
      Contact( #St_Opening )
   END_RUNG wire#w1
   RUNG wire#powerrail
      Contact( #FbClosed )
      wire#w2
      Coil( #Close_Reached )
   END_RUNG
   RUNG wire#powerrail
      Contact( #TON_Move.Q )
      Contact( #St_Closing )
   END_RUNG wire#w2
   // the same network as SCL:
   #Open_Reached := #FbOpen OR (#TON_Move.Q AND #St_Opening);
   #Close_Reached := #FbClosed OR (#TON_Move.Q AND #St_Closing);
END_REGION

REGION Network 10: Drive coils (works for 1‑coil and 2‑coil valves)
   // Two‑coil: energize Q_Open only while opening and Q_Close only while closing (spool stays latched).
   // One‑coil: energize Q_Open continuously whenever the final desired state is Open and no faults; de‑energize to close.
   RUNG wire#powerrail
      Contact( #St_Opening )
      Contact( #TwoCoils )
      wire#w1
      Coil( #Q_Open )
   END_RUNG
   RUNG wire#powerrail
      I_Contact( #TwoCoils )
      Contact( #Cmd_DesiredOpen_OK )
      I_Contact( #FaultTO )
      I_Contact( #FaultFB )
      I_Contact( #OOS )
      Contact( #Permissive )
   END_RUNG wire#w1
   RUNG wire#powerrail
      Contact( #St_Closing )
      Contact( #TwoCoils )
      Coil( #Q_Close )
   END_RUNG
   // the same network as SCL:
   #Q_Open := (#St_Opening AND #TwoCoils) OR (NOT #TwoCoils AND #Cmd_DesiredOpen_OK AND NOT #FaultTO AND NOT #FaultFB AND NOT #OOS AND #Permissive);
   #Q_Close := #St_Closing AND #TwoCoils;
END_REGION

REGION Network 11: Ready flag
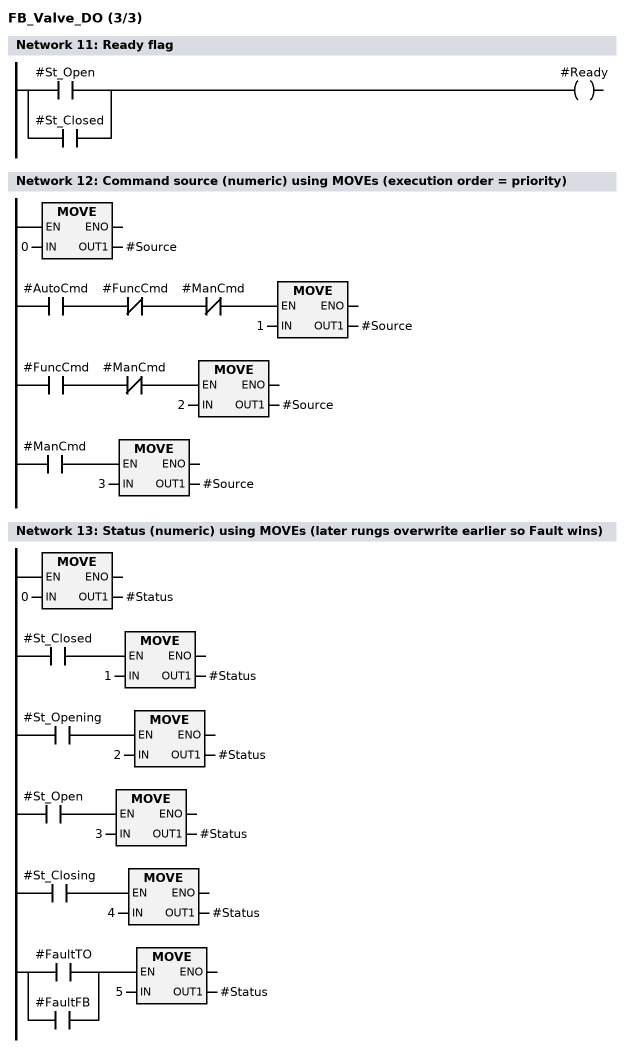
   RUNG wire#powerrail
      Contact( #St_Open )
      wire#w1
      Coil( #Ready )
   END_RUNG
   RUNG wire#powerrail
      Contact( #St_Closed )
   END_RUNG wire#w1
   // the same network as SCL:
   #Ready := #St_Open OR #St_Closed;
END_REGION

REGION Network 12: Command source (numeric) using MOVEs (execution order = priority)
   RUNG wire#powerrail
      Move(in := 0, out1 => #Source)
   END_RUNG
   RUNG wire#powerrail
      Contact( #AutoCmd )
      I_Contact( #FuncCmd )
      I_Contact( #ManCmd )
      Move(in := 1, out1 => #Source)
   END_RUNG
   RUNG wire#powerrail
      Contact( #FuncCmd )
      I_Contact( #ManCmd )
      Move(in := 2, out1 => #Source)
   END_RUNG
   RUNG wire#powerrail
      Contact( #ManCmd )
      Move(in := 3, out1 => #Source)
   END_RUNG
   // the same network as SCL:
   #Source := 0;
   IF #AutoCmd AND NOT #FuncCmd AND NOT #ManCmd THEN #Source := 1; END_IF;
   IF #FuncCmd AND NOT #ManCmd THEN #Source := 2; END_IF;
   IF #ManCmd THEN #Source := 3; END_IF;
END_REGION

REGION Network 13: Status (numeric) using MOVEs (later rungs overwrite earlier so Fault wins)
   RUNG wire#powerrail
      Move(in := 0, out1 => #Status)
   END_RUNG
   RUNG wire#powerrail
      Contact( #St_Closed )
      Move(in := 1, out1 => #Status)
   END_RUNG
   RUNG wire#powerrail
      Contact( #St_Opening )
      Move(in := 2, out1 => #Status)
   END_RUNG
   RUNG wire#powerrail
      Contact( #St_Open )
      Move(in := 3, out1 => #Status)
   END_RUNG
   RUNG wire#powerrail
      Contact( #St_Closing )
      Move(in := 4, out1 => #Status)
   END_RUNG
   RUNG wire#powerrail
      Contact( #FaultTO )
      wire#w1
      Move(in := 5, out1 => #Status)
   END_RUNG
   RUNG wire#powerrail
      Contact( #FaultFB )
   END_RUNG wire#w1
   // the same network as SCL:
   #Status := 0;
   IF #St_Closed THEN #Status := 1; END_IF;
   IF #St_Opening THEN #Status := 2; END_IF;
   IF #St_Open THEN #Status := 3; END_IF;
   IF #St_Closing THEN #Status := 4; END_IF;
   IF #FaultTO OR #FaultFB THEN #Status := 5; END_IF;
END_REGION
END_FUNCTION_BLOCK

FUNCTION_BLOCK "FB_Motor_VFD"   // FB2, LAD
{ S7_Optimized_Access := 'TRUE' }
VERSION : 0.1
   VAR_INPUT
      Start_Auto : Bool;
      Start_Func : Bool;
      Start_Man : Bool;
      OOS : Bool;
      RevDwell : Time := T#2S;
      Permissive : Bool := true;
      PulseEnable : Bool;   // TRUE = do Fwd/Hold/Bwd pulsing
      T_Fwd : Time := T#8S;
      T_Hold : Time := T#2S;
      T_Bwd : Time := T#6S;
      DischargeMode : Bool;   // TRUE = forward only
      SpeedSP_pct : Real;   // 0..100, normal speed
      DischSpeed_pct : Real;   // 0..100, used when DischargeMode=TRUE
      DriveReady : Bool;   // optional, from VFD
      DriveFault : Bool;   // optional, from VFD
      StartTimeout : Time := T#5S;
   END_VAR
   VAR_OUTPUT
      Q_Run : Bool;   // to RUN relay or PN run bit
      Q_DirFwd : Bool;   // TRUE = forward, FALSE = reverse
      AO_SpeedPct : Real;   // speed command 0..100%
      Running : Bool;
      Direction : UInt;   // 0 Stop, 1 Fwd, 2 Bwd
      Fault : Bool;
      FaultCode : UInt;   // 0 ok, 1 timeout, 2 drive fault, 3 permissive/OOS
      Source : UInt;   // 1 Auto, 2 Func, 3 Man
      R_Fwd : Bool;
      R_Rev : Bool;
      State : UInt;   // 0 Stop, 1 Fwd, 2 Hold, 3 Bwd (for HMI)
      RDwell_Q : Bool;
   END_VAR
   VAR
      Start_Prio : Bool;
      RunCmd : Bool;
      Start_OK : Bool;
      RStart : R_TRIG;
      St_Fwd : Bool;
      St_Hold : Bool;
      St_Bwd : Bool;
      Tmr_Fwd : TON_TIME;
      Tmr_Hold : TON_TIME;
      Tmr_Bwd : TON_TIME;
      Tmr_Dwell : TON_TIME;
      DwellActive : Bool;
      PrevDirFwd : Bool;
      Tmr_Start : TON_TIME;
      StartRise : Bool;
      PulseActive : Bool;
      RDwell : R_TRIG;
      FDwell : F_TRIG;
      ChangePulse : Bool;
      DwellRun : Bool;
      Start_Raw : Bool;
      DirFwdCmd : Bool;
   END_VAR
BEGIN

REGION Network 1: Command priority (Man > Func > Auto) → Start_Raw
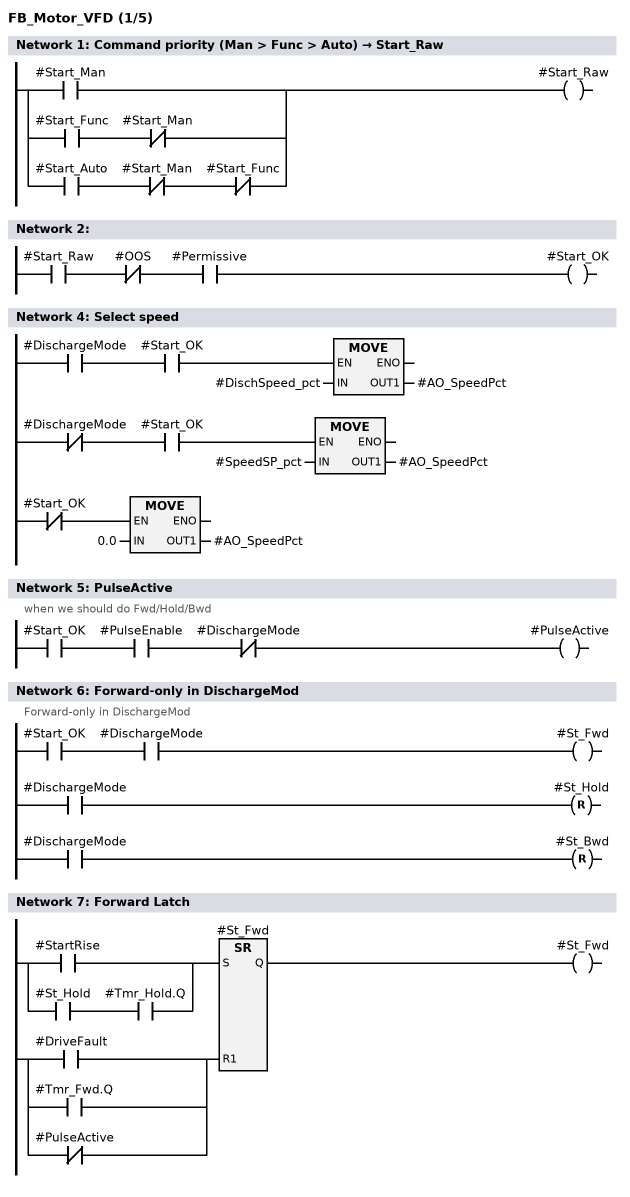
   RUNG wire#powerrail
      Contact( #Start_Man )
      wire#w1
      Coil( #Start_Raw )
   END_RUNG
   RUNG wire#powerrail
      Contact( #Start_Func )
      I_Contact( #Start_Man )
   END_RUNG wire#w1
   RUNG wire#powerrail
      Contact( #Start_Auto )
      I_Contact( #Start_Man )
      I_Contact( #Start_Func )
   END_RUNG wire#w1
   // the same network as SCL:
   #Start_Raw := #Start_Man OR (#Start_Func AND NOT #Start_Man) OR (#Start_Auto AND NOT #Start_Man AND NOT #Start_Func);
END_REGION

REGION Network 2
   RUNG wire#powerrail
      Contact( #Start_Raw )
      I_Contact( #OOS )
      Contact( #Permissive )
      Coil( #Start_OK )
   END_RUNG
   // the same network as SCL:
   #Start_OK := #Start_Raw AND NOT #OOS AND #Permissive;
END_REGION

REGION Network 3 (SCL)
   // CORRECT:
   #RStart(CLK := #Start_OK);
   #StartRise := #RStart.Q;
END_REGION

REGION Network 4: Select speed
   RUNG wire#powerrail
      Contact( #DischargeMode )
      Contact( #Start_OK )
      Move(in := #DischSpeed_pct, out1 => #AO_SpeedPct)
   END_RUNG
   RUNG wire#powerrail
      I_Contact( #DischargeMode )
      Contact( #Start_OK )
      Move(in := #SpeedSP_pct, out1 => #AO_SpeedPct)
   END_RUNG
   RUNG wire#powerrail
      I_Contact( #Start_OK )
      Move(in := 0.0, out1 => #AO_SpeedPct)
   END_RUNG
   // the same network as SCL:
   IF #DischargeMode AND #Start_OK THEN #AO_SpeedPct := #DischSpeed_pct; END_IF;
   IF NOT #DischargeMode AND #Start_OK THEN #AO_SpeedPct := #SpeedSP_pct; END_IF;
   IF NOT #Start_OK THEN #AO_SpeedPct := 0.0; END_IF;
END_REGION

REGION Network 5: PulseActive
   // when we should do Fwd/Hold/Bwd
   RUNG wire#powerrail
      Contact( #Start_OK )
      Contact( #PulseEnable )
      I_Contact( #DischargeMode )
      Coil( #PulseActive )
   END_RUNG
   // the same network as SCL:
   #PulseActive := #Start_OK AND #PulseEnable AND NOT #DischargeMode;
END_REGION

REGION Network 6: Forward-only in DischargeMod
   // Forward-only in DischargeMod
   RUNG wire#powerrail
      Contact( #Start_OK )
      Contact( #DischargeMode )
      Coil( #St_Fwd )
   END_RUNG
   RUNG wire#powerrail
      Contact( #DischargeMode )
      R_Coil( #St_Hold )
   END_RUNG
   RUNG wire#powerrail
      Contact( #DischargeMode )
      R_Coil( #St_Bwd )
   END_RUNG
   // the same network as SCL:
   #St_Fwd := #Start_OK AND #DischargeMode;
   IF #DischargeMode THEN
       #St_Hold := FALSE;
       #St_Bwd := FALSE;
   END_IF;
END_REGION

REGION Network 7: Forward Latch
   RUNG wire#powerrail
      Contact( #StartRise )
      wire#w1
      S_SR(operand := #St_Fwd, r1 := wire#w2)
      Coil( #St_Fwd )
   END_RUNG
   RUNG wire#powerrail
      Contact( #St_Hold )
      Contact( #Tmr_Hold.Q )
   END_RUNG wire#w1
   RUNG wire#powerrail
      Contact( #DriveFault )
   END_RUNG wire#w2
   RUNG wire#powerrail
      Contact( #Tmr_Fwd.Q )
   END_RUNG wire#w2
   RUNG wire#powerrail
      I_Contact( #PulseActive )
   END_RUNG wire#w2
   // the same network as SCL:
   IF #StartRise OR (#St_Hold AND #Tmr_Hold.Q) THEN
       #St_Fwd := TRUE;   // SR flip-flop
   END_IF;
   IF #DriveFault OR #Tmr_Fwd.Q OR NOT #PulseActive THEN #St_Fwd := FALSE; END_IF;
   #St_Fwd := #St_Fwd;
END_REGION

REGION Network 8: Hold Latch
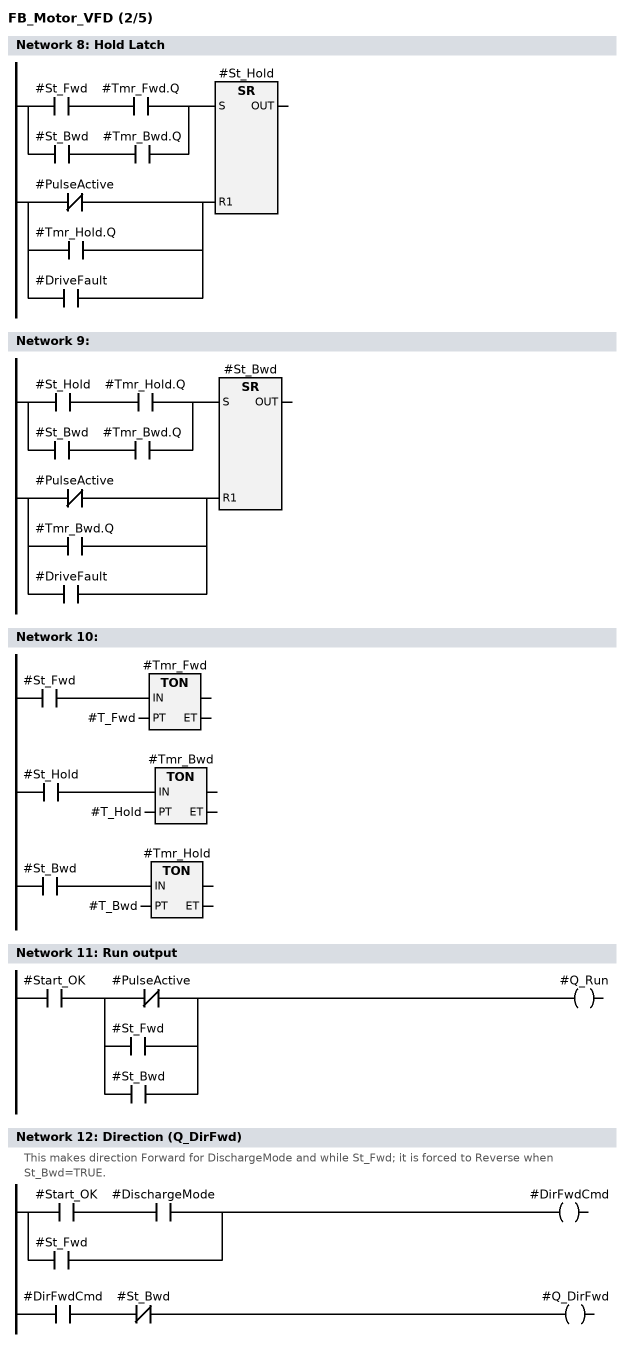
   RUNG wire#powerrail
      Contact( #St_Fwd )
      Contact( #Tmr_Fwd.Q )
      wire#w1
      S_SR(operand := #St_Hold, r1 := wire#w2)
   END_RUNG
   RUNG wire#powerrail
      Contact( #St_Bwd )
      Contact( #Tmr_Bwd.Q )
   END_RUNG wire#w1
   RUNG wire#powerrail
      I_Contact( #PulseActive )
   END_RUNG wire#w2
   RUNG wire#powerrail
      Contact( #Tmr_Hold.Q )
   END_RUNG wire#w2
   RUNG wire#powerrail
      Contact( #DriveFault )
   END_RUNG wire#w2
   // the same network as SCL:
   IF (#St_Fwd AND #Tmr_Fwd.Q) OR (#St_Bwd AND #Tmr_Bwd.Q) THEN
       #St_Hold := TRUE;   // SR flip-flop
   END_IF;
   IF NOT #PulseActive OR #Tmr_Hold.Q OR #DriveFault THEN #St_Hold := FALSE; END_IF;
END_REGION

REGION Network 9
   RUNG wire#powerrail
      Contact( #St_Hold )
      Contact( #Tmr_Hold.Q )
      wire#w1
      S_SR(operand := #St_Bwd, r1 := wire#w2)
   END_RUNG
   RUNG wire#powerrail
      Contact( #St_Bwd )
      Contact( #Tmr_Bwd.Q )
   END_RUNG wire#w1
   RUNG wire#powerrail
      I_Contact( #PulseActive )
   END_RUNG wire#w2
   RUNG wire#powerrail
      Contact( #Tmr_Bwd.Q )
   END_RUNG wire#w2
   RUNG wire#powerrail
      Contact( #DriveFault )
   END_RUNG wire#w2
   // the same network as SCL:
   IF (#St_Hold AND #Tmr_Hold.Q) OR (#St_Bwd AND #Tmr_Bwd.Q) THEN
       #St_Bwd := TRUE;   // SR flip-flop
   END_IF;
   IF NOT #PulseActive OR #Tmr_Bwd.Q OR #DriveFault THEN #St_Bwd := FALSE; END_IF;
END_REGION

REGION Network 10
   #Tmr_Fwd(IN := #St_Fwd, PT := #T_Fwd);   // TON
   #Tmr_Bwd(IN := #St_Hold, PT := #T_Hold);   // TON
   #Tmr_Hold(IN := #St_Bwd, PT := #T_Bwd);   // TON
END_REGION

REGION Network 11: Run output
   RUNG wire#powerrail
      Contact( #Start_OK )
      wire#w1
      I_Contact( #PulseActive )
      wire#w2
      Coil( #Q_Run )
   END_RUNG
   RUNG wire#w1
      Contact( #St_Fwd )
   END_RUNG wire#w2
   RUNG wire#w1
      Contact( #St_Bwd )
   END_RUNG wire#w2
   // the same network as SCL:
   #Q_Run := #Start_OK AND (NOT #PulseActive OR #St_Fwd OR #St_Bwd);
END_REGION

REGION Network 12: Direction (Q_DirFwd)
   // This makes direction Forward for DischargeMode and while St_Fwd; it is forced to Reverse when St_Bwd=TRUE.
   RUNG wire#powerrail
      Contact( #Start_OK )
      Contact( #DischargeMode )
      wire#w1
      Coil( #DirFwdCmd )
   END_RUNG
   RUNG wire#powerrail
      Contact( #St_Fwd )
   END_RUNG wire#w1
   RUNG wire#powerrail
      Contact( #DirFwdCmd )
      I_Contact( #St_Bwd )
      Coil( #Q_DirFwd )
   END_RUNG
   // the same network as SCL:
   #DirFwdCmd := (#Start_OK AND #DischargeMode) OR #St_Fwd;
   #Q_DirFwd := #DirFwdCmd AND NOT #St_Bwd;
END_REGION

REGION Network 13: Detect change of direction
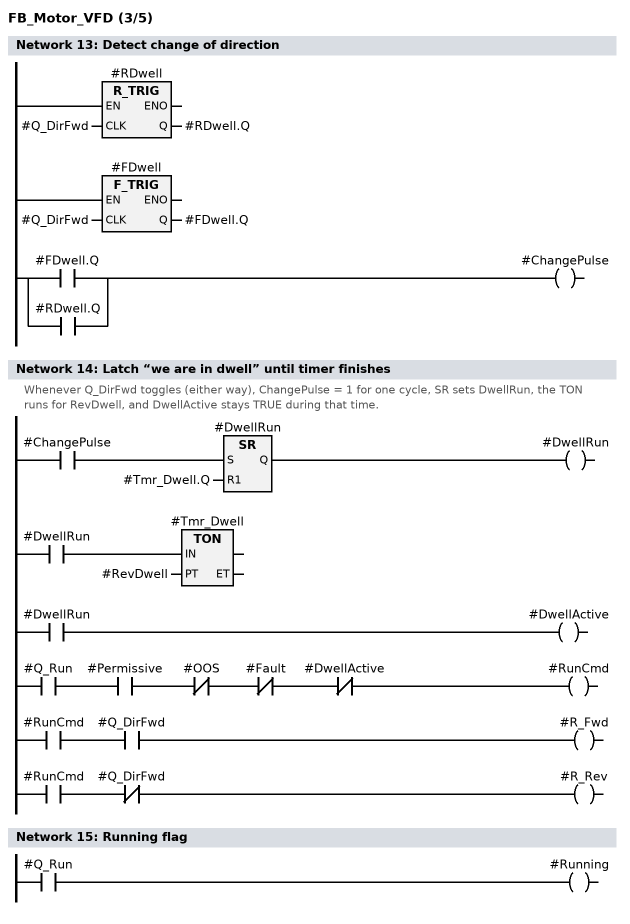
   #RDwell(CLK := #Q_DirFwd, Q => #RDwell.Q);   // R_TRIG
   #FDwell(CLK := #Q_DirFwd, Q => #FDwell.Q);   // F_TRIG
   #ChangePulse := #FDwell.Q OR #RDwell.Q;
END_REGION

REGION Network 14: Latch “we are in dwell” until timer finishes
   // Whenever Q_DirFwd toggles (either way), ChangePulse = 1 for one cycle, SR sets DwellRun, the TON runs for RevDwell, and DwellActive stays TRUE during that time.
   IF #ChangePulse THEN
       #DwellRun := TRUE;   // SR flip-flop
   END_IF;
   IF #Tmr_Dwell.Q THEN #DwellRun := FALSE; END_IF;
   #DwellRun := #DwellRun;
   #Tmr_Dwell(IN := #DwellRun, PT := #RevDwell);   // TON
   #DwellActive := #DwellRun;
   #RunCmd := #Q_Run AND #Permissive AND NOT #OOS AND NOT #Fault AND NOT #DwellActive;
   #R_Fwd := #RunCmd AND #Q_DirFwd;
   #R_Rev := #RunCmd AND NOT #Q_DirFwd;
END_REGION

REGION Network 15: Running flag
   RUNG wire#powerrail
      Contact( #Q_Run )
      Coil( #Running )
   END_RUNG
   // the same network as SCL:
   #Running := #Q_Run;
END_REGION

REGION Network 16: Start timeout and Drive faults
   // if you don’t have DriveReady wiring yet, set DriveReady=TRUE when you CALL the FB so the start timeout won’t trigger.
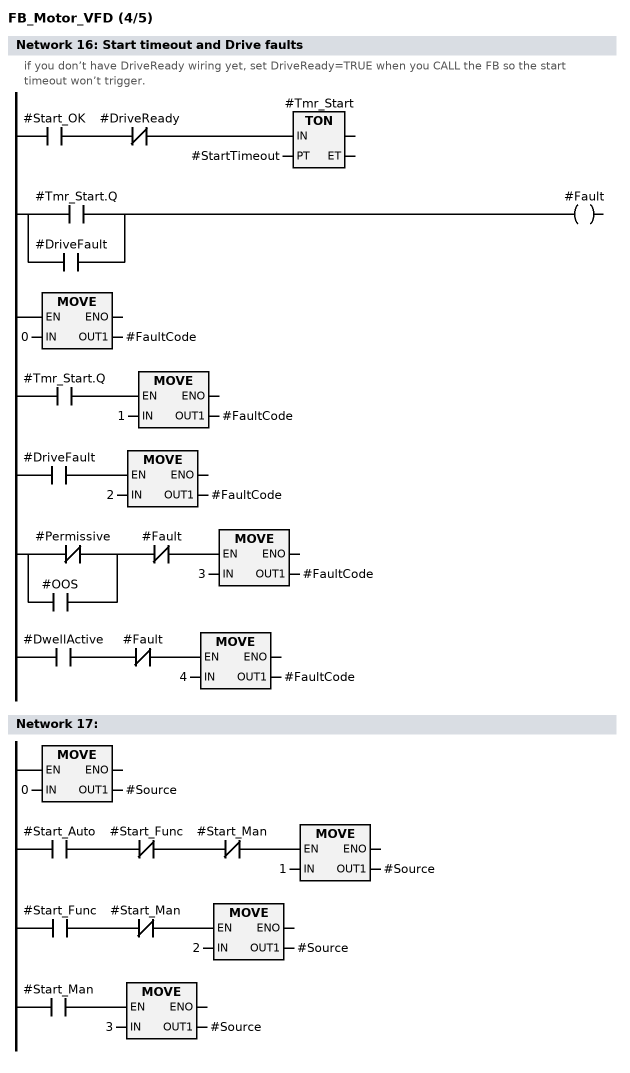
   #Tmr_Start(IN := #Start_OK AND NOT #DriveReady, PT := #StartTimeout);   // TON
   #Fault := #Tmr_Start.Q OR #DriveFault;
   #FaultCode := 0;
   IF #Tmr_Start.Q THEN #FaultCode := 1; END_IF;
   IF #DriveFault THEN #FaultCode := 2; END_IF;
   IF (NOT #Permissive OR #OOS) AND NOT #Fault THEN #FaultCode := 3; END_IF;
   IF #DwellActive AND NOT #Fault THEN #FaultCode := 4; END_IF;
END_REGION

REGION Network 17
   RUNG wire#powerrail
      Move(in := 0, out1 => #Source)
   END_RUNG
   RUNG wire#powerrail
      Contact( #Start_Auto )
      I_Contact( #Start_Func )
      I_Contact( #Start_Man )
      Move(in := 1, out1 => #Source)
   END_RUNG
   RUNG wire#powerrail
      Contact( #Start_Func )
      I_Contact( #Start_Man )
      Move(in := 2, out1 => #Source)
   END_RUNG
   RUNG wire#powerrail
      Contact( #Start_Man )
      Move(in := 3, out1 => #Source)
   END_RUNG
   // the same network as SCL:
   #Source := 0;
   IF #Start_Auto AND NOT #Start_Func AND NOT #Start_Man THEN #Source := 1; END_IF;
   IF #Start_Func AND NOT #Start_Man THEN #Source := 2; END_IF;
   IF #Start_Man THEN #Source := 3; END_IF;
END_REGION

REGION Network 18: State
   // for HMI: 0 Stop, 1 Fwd, 2 Hold, 3 Bwd
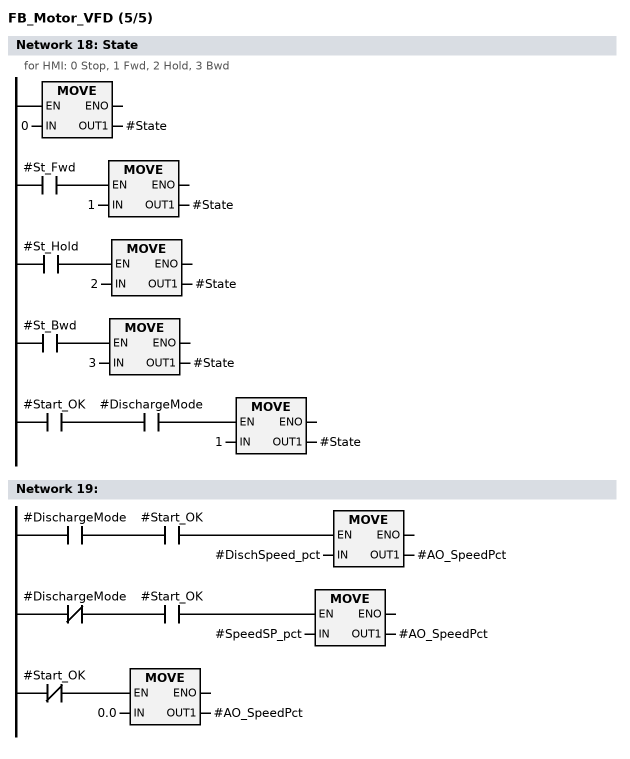
   RUNG wire#powerrail
      Move(in := 0, out1 => #State)
   END_RUNG
   RUNG wire#powerrail
      Contact( #St_Fwd )
      Move(in := 1, out1 => #State)
   END_RUNG
   RUNG wire#powerrail
      Contact( #St_Hold )
      Move(in := 2, out1 => #State)
   END_RUNG
   RUNG wire#powerrail
      Contact( #St_Bwd )
      Move(in := 3, out1 => #State)
   END_RUNG
   RUNG wire#powerrail
      Contact( #Start_OK )
      Contact( #DischargeMode )
      Move(in := 1, out1 => #State)
   END_RUNG
   // the same network as SCL:
   #State := 0;
   IF #St_Fwd THEN #State := 1; END_IF;
   IF #St_Hold THEN #State := 2; END_IF;
   IF #St_Bwd THEN #State := 3; END_IF;
   IF #Start_OK AND #DischargeMode THEN #State := 1; END_IF;
END_REGION

REGION Network 19
   RUNG wire#powerrail
      Contact( #DischargeMode )
      Contact( #Start_OK )
      Move(in := #DischSpeed_pct, out1 => #AO_SpeedPct)
   END_RUNG
   RUNG wire#powerrail
      I_Contact( #DischargeMode )
      Contact( #Start_OK )
      Move(in := #SpeedSP_pct, out1 => #AO_SpeedPct)
   END_RUNG
   RUNG wire#powerrail
      I_Contact( #Start_OK )
      Move(in := 0.0, out1 => #AO_SpeedPct)
   END_RUNG
   // the same network as SCL:
   IF #DischargeMode AND #Start_OK THEN #AO_SpeedPct := #DischSpeed_pct; END_IF;
   IF NOT #DischargeMode AND #Start_OK THEN #AO_SpeedPct := #SpeedSP_pct; END_IF;
   IF NOT #Start_OK THEN #AO_SpeedPct := 0.0; END_IF;
END_REGION
END_FUNCTION_BLOCK

FUNCTION_BLOCK "FB_Motor_Controller"   // FB4, SCL
{ S7_Optimized_Access := 'TRUE' }
VERSION : 0.1
   VAR_INPUT
      Enable : Bool;
      Command_Start : Bool;
      Command_Stop : Bool;
      Speed_Setpoint : Real;
      Pulse_Enable : Bool;
      Discharge_Mode : Bool;
      Direction_Command : Int;
      Safety_Permissive : Bool;
      Reset_Command : Bool;
   END_VAR
   VAR_OUTPUT
      Motor_Running : Bool;
      Motor_Ready : Bool;
      Motor_Fault : Bool;
      Current_Speed : Real;
      Current_Direction : UInt;
      Status_Text : String;
      Direction : UInt;
   END_VAR
   VAR_IN_OUT
      Motor_FB : "FB_Motor_VFD";
   END_VAR
   VAR
      Speed_Ramp_Timer : TON_TIME;
      Direction_Timer : TON_TIME;
      Target_Speed : Real;
      Direction_Change : Bool;
      Previous_Direction : Int;
   END_VAR
BEGIN
   // Update motor 1 data directly in DB
   "DB_Motors".Motors[1].Config.Motor_Name := 'SCREW_MOTOR';
   "DB_Motors".Motors[1].Interlocks.Permissive := #Safety_Permissive;
   "DB_Motors".Motors[1].Interlocks.OOS := NOT #Enable;
   // Speed ramping
   IF #Enable AND #Safety_Permissive THEN
       IF ABS(#Speed_Setpoint - #Target_Speed) > 1.0 THEN
           #Speed_Ramp_Timer(IN := TRUE,
                             PT := T#100MS);
           IF #Speed_Ramp_Timer.Q THEN
               IF #Speed_Setpoint > #Target_Speed THEN
                   #Target_Speed := #Target_Speed + 2.0;
               ELSE
                   #Target_Speed := #Target_Speed - 2.0;
               END_IF;
               #Speed_Ramp_Timer(IN := FALSE,
                                 PT := T#0S);
           END_IF;
       ELSE
           #Target_Speed := #Speed_Setpoint;
       END_IF;

       // Set commands in DB
       "DB_Motors".Motors[1].Command.Start_Auto := #Command_Start;
       "DB_Motors".Motors[1].Command.Speed_SP_pct := #Target_Speed;
       "DB_Motors".Motors[1].Command.Pulse_Enable := #Pulse_Enable;
       "DB_Motors".Motors[1].Command.Discharge_Mode := #Discharge_Mode;
       "DB_Motors".Motors[1].Command.Direction := #Direction_Command;
   ELSE
       "DB_Motors".Motors[1].Command.Start_Auto := FALSE;
       "DB_Motors".Motors[1].Command.Speed_SP_pct := 0.0;
       #Target_Speed := 0.0;
   END_IF;
   // Call YOUR FB_Motor_VFD
   #Motor_FB(
             Start_Auto := "DB_Motors".Motors[1].Command.Start_Auto,
             Start_Func := "DB_Motors".Motors[1].Command.Start_Func,
             Start_Man := "DB_Motors".Motors[1].Command.Start_Man,
             OOS := "DB_Motors".Motors[1].Interlocks.OOS,
             RevDwell := "DB_Motors".Motors[1].Config.Rev_Dwell,
             Permissive := "DB_Motors".Motors[1].Interlocks.Permissive,
             PulseEnable := "DB_Motors".Motors[1].Command.Pulse_Enable,
             T_Fwd := "DB_Motors".Motors[1].Config.T_Fwd,
             T_Hold := "DB_Motors".Motors[1].Config.T_Hold,
             T_Bwd := "DB_Motors".Motors[1].Config.T_Bwd,
             DischargeMode := "DB_Motors".Motors[1].Command.Discharge_Mode,
             SpeedSP_pct := "DB_Motors".Motors[1].Command.Speed_SP_pct,
             DischSpeed_pct := "DB_Motors".Motors[1].Config.Disch_Speed_pct,
             DriveReady := TRUE,
             DriveFault := FALSE,
             StartTimeout := "DB_Motors".Motors[1].Config.Start_Timeout,

             Q_Run => "DB_Motors".Motors[1].Outputs.Q_Run,
             Q_DirFwd => "DB_Motors".Motors[1].Outputs.Q_DirFwd,
             AO_SpeedPct => "DB_Motors".Motors[1].Outputs.AO_SpeedPct,
             Running => "DB_Motors".Motors[1].Status.Running,
             Direction => "DB_Motors".Motors[1].Status.Direction,
             Fault => "DB_Motors".Motors[1].Status.Fault,
             Source => "DB_Motors".Motors[1].Status.Source,
             State => "DB_Motors".Motors[1].Status.State
   );
   // Outputs
   #Motor_Running := "DB_Motors".Motors[1].Status.Running;
   #Motor_Ready := "DB_Motors".Motors[1].Interlocks.Permissive AND NOT "DB_Motors".Motors[1].Status.Fault;
   #Motor_Fault := "DB_Motors".Motors[1].Status.Fault;
   #Current_Speed := "DB_Motors".Motors[1].Outputs.AO_SpeedPct;

   IF #Motor_Fault THEN
       #Status_Text := 'Motor fault active';
   ELSIF #Motor_Running THEN
       #Status_Text := 'Motor running';
   ELSE
       #Status_Text := 'Motor stopped';
   END_IF;
END_FUNCTION_BLOCK

FUNCTION_BLOCK "FB_Preparation_Phase"   // FB5, SCL
{ S7_Optimized_Access := 'TRUE' }
VERSION : 0.1
   VAR_INPUT
      Phase_Enable : Bool;
      Safety_Permissive : Bool;
      Reset_Phase : Bool;
   END_VAR
   VAR_OUTPUT
      Phase_Complete : Bool;
      Phase_Active : Bool;
      Phase_Fault : Bool;
      Step_Complete : Bool;
      Phase_Status : String;
      Step_Status : String;
      Phase_Progress : Real;
      Next_Step : UInt;
   END_VAR
   VAR_IN_OUT
      Current_Step : UInt;
   END_VAR
   VAR
      Phase_Timers : Array[1..10] of TON_TIME;
      Total_Steps : UInt := 5;
      Completed_Steps : UInt;
      Step_Complete_15 : Bool;
      Step_Complete_1 : Bool;
      Step_Complete_2 : Bool;
      Step_Complete_3 : Bool;
      Step_Complete_4 : Bool;
      Step_Fault_Flag : Bool;
      Timer_Step_15 : TON_TIME;
      Time_text1 : TON_TIME;
      Timer_Step_1 : TON_TIME;
      Timer_Step_2 : TON_TIME;
      Timer_Step_3 : TON_TIME;
      Timer_Step_4 : TON_TIME;
   END_VAR
   VAR_TEMP
      i : Int;
      Temp_Step_Active : Bool;
      Temp_Fault_Code : UInt;
      Temp_Time_Remaining : Time;
      Temp_Water_Added : Real;
      Temp_Wait_Time : Time;
   END_VAR
BEGIN
   #Phase_Fault := FALSE;

   IF #Reset_Phase THEN
       #Phase_Complete := FALSE;
       #Phase_Active := FALSE;
       #Phase_Fault := FALSE;
       #Step_Complete := FALSE;
       #Current_Step := 15;
       #Phase_Status := 'Phase reset';
       #Phase_Progress := 0.0;
       #Completed_Steps := 0;
       RETURN;
   END_IF;

   IF #Phase_Enable AND #Safety_Permissive THEN
       #Phase_Active := TRUE;
       #Phase_Status := 'Preparation phase active';

       CASE #Current_Step OF
           15: // Lock Discharge Door
               "FC_Lock_Discharge_Door"(
                                        Step_Enable := TRUE,
                                        Safety_OK := #Safety_Permissive,
                                        Step_Timeout := T#30S,
                                        Door_Locked_FB := "DB_Process".IO.Door_Locked_FB,
                                        Reset_Step := "DB_Process".HMI.Reset_p_s,
                                        Close_Timer:=#Phase_Timers[1],
                                        Step_Timer := #Timer_Step_15,
                                        Step_Complete => #Step_Complete,
                                        Step_Active => #Temp_Step_Active,        // ✅ ASSIGN TO TEMP
                                        Step_Fault => #Step_Fault_Flag,
                                        Fault_Code => #Temp_Fault_Code,          // ✅ ASSIGN TO TEMP
                                        Status_Text => #Step_Status,
                                        Time_Remaining => #Temp_Time_Remaining   // ✅ ASSIGN TO TEMP
               );

               IF #Step_Complete THEN
                   #Next_Step := 1;
                   #Current_Step := #Next_Step;
                   #Completed_Steps := 1;
               END_IF;

           1: // Add Water
               "FC_Add_Water"(
                              Step_Enable := TRUE,
                              Safety_OK := #Safety_Permissive,
                              Step_Timeout := "DB_Recipes".Active_Recipe.Production.Water_Flow_Timeout,
                              Water_Level_FB => "DB_Process".IO.Water_Level_FB,
                              Target_Quantity := "DB_Recipes".Active_Recipe.Production.Adding_Water1_QTY,
                              Flow_Rate := "DB_Process".IO.AI_Water_Flow,
                              Reset_Step := "DB_Process".HMI.Reset_p_s,

                              Step_Timer := #Timer_Step_1,

                              Step_Complete => #Step_Complete,
                              Step_Active => #Temp_Step_Active,        // ✅ ASSIGN TO TEMP
                              Step_Fault => #Step_Fault_Flag,
                              Fault_Code => #Temp_Fault_Code,          // ✅ ASSIGN TO TEMP
                              Status_Text => #Step_Status,
                              Water_Added => #Temp_Water_Added,        // ✅ ASSIGN TO TEMP
                              Time_Remaining => #Temp_Time_Remaining   // ✅ ASSIGN TO TEMP
               );
               "DB_Process".Status.Water_Level_Actual := #Temp_Water_Added;

               IF #Step_Complete THEN
                   #Next_Step := 2;
                   #Current_Step := #Next_Step;
                   #Completed_Steps := 2;
               END_IF;

           2: // Open Manhole /add timer to show the status
               "FC_Open_Manhole"(
                                 Step_Enable := TRUE,
                                 Safety_OK := #Safety_Permissive,
                                 Step_Timeout := "DB_Recipes".Active_Recipe.Production.Manhole_Open_Time,
                                 Manhole_Open_FB := "DB_Process".IO.Manhole_Open_FB,
                                 Manhole_Closed_FB := "DB_Process".IO.Manhole_Closed_FB,
                                 Reset_Step := "DB_Process".HMI.Reset_p_s,

                                 Step_Timer := #Timer_Step_2,
                                 Open_Timer:=#Phase_Timers[2],
                                 Step_Complete => #Step_Complete,
                                 Step_Active => #Temp_Step_Active,        // ✅ ASSIGN TO TEMP
                                 Step_Fault => #Step_Fault_Flag,
                                 Fault_Code => #Temp_Fault_Code,          // ✅ ASSIGN TO TEMP
                                 Status_Text => #Step_Status,
                                 Time_Remaining => #Temp_Time_Remaining   // ✅ ASSIGN TO TEMP
               );

               IF #Step_Complete THEN
                   #Next_Step := 3;
                   #Current_Step := #Next_Step;
                   #Completed_Steps := 3;
               END_IF;

           3: // Wait for Raw Materials  
               "FC_Wait_Raw_Materials"(
                                       Step_Enable := TRUE,
                                       Safety_OK := #Safety_Permissive,
                                       RawMat_Confirm := "DB_Process".HMI.RawMaterial_OK,
                                       Manhole_Open_FB := "DB_Process".IO.Manhole_Open_FB,
                                       Manhole_Closed_FB := "DB_Process".IO.Manhole_Closed_FB,
                                       Max_Wait_Time := T#30S,
                                       Reset_Step := "DB_Process".HMI.Reset_p_s,

                                       Wait_Timer := #Timer_Step_3,

                                       Step_Complete => #Step_Complete,
                                       Step_Active => #Temp_Step_Active,        // ✅ ASSIGN TO TEMP
                                       Step_Fault => #Step_Fault_Flag,
                                       Fault_Code => #Temp_Fault_Code,          // ✅ ASSIGN TO TEMP
                                       Status_Text => #Step_Status,
                                       Wait_Time_Elapsed => #Temp_Wait_Time     // ✅ ASSIGN TO TEMP
               );

               IF #Step_Complete THEN
                   #Next_Step := 4;
                   #Current_Step := #Next_Step;
                   #Completed_Steps := 4;
               END_IF;

           4: // Close Manhole add timer to show the status
               "FC_Close_Manhole"(
                                  Step_Enable := TRUE,
                                  Safety_OK := #Safety_Permissive,
                                  Step_Timeout := "DB_Recipes".Active_Recipe.Production.Manhole_Close_Time,
                                  Manhole_Closed_FB := "DB_Process".IO.Manhole_Closed_FB,
                                  Manhole_Open_FB := "DB_Process".IO.Manhole_Open_FB,
                                  Reset_Step := "DB_Process".HMI.Reset_p_s,

                                  Step_Timer := #Timer_Step_4,
                                  Close_Timer:=#Phase_Timers[3],
                                  Step_Complete => #Step_Complete,
                                  Step_Active => #Temp_Step_Active,        // ✅ ASSIGN TO TEMP
                                  Step_Fault => #Step_Fault_Flag,
                                  Fault_Code => #Temp_Fault_Code,          // ✅ ASSIGN TO TEMP
                                  Status_Text => #Step_Status,
                                  Time_Remaining => #Temp_Time_Remaining   // ✅ ASSIGN TO TEMP
               );

               IF #Step_Complete THEN
                   #Phase_Complete := TRUE;
                   #Next_Step := 5;
                   #Current_Step := #Next_Step;
                   #Completed_Steps := 5;
                   #Phase_Status := 'Preparation complete';
               END_IF;

           ELSE
               #Phase_Fault := TRUE;
               #Phase_Status := 'Invalid step';
       END_CASE;

       #Phase_Progress := (UINT_TO_REAL(#Completed_Steps) / UINT_TO_REAL(#Total_Steps)) * 100.0;

   ELSE
       #Phase_Active := FALSE;
       #Phase_Complete := FALSE;
       #Phase_Status := 'Phase disabled';
   END_IF;
END_FUNCTION_BLOCK

FUNCTION_BLOCK "FB_Temperature_Controller"   // FB6, SCL
{ S7_Optimized_Access := 'TRUE' }
VERSION : 0.1
   VAR_INPUT
      Enable_Control : Bool;
      Temperature_SP : Real;
      Temperature_PV : Real;
      Control_Deadband : Real;
      Safety_Permissive : Bool;
   END_VAR
   VAR_OUTPUT
      Control_Active : Bool;
      At_Setpoint : Bool;
      Heating_Active : Bool;
      Cooling_Active : Bool;
      Status_Text : String;
      Temp_Error : Real;
   END_VAR
   VAR
      Control_Timer : TON_TIME;
      Setpoint_Active : Real;
      High_Limit : Real := 100.0;
      Low_Limit : Real := 0.0;
      Control_Cycle : Time := T#2S;
      Enable_Internal : Bool;
   END_VAR
BEGIN
   #Heating_Active := FALSE;
   #Cooling_Active := FALSE;

   IF #Enable_Control AND #Safety_Permissive THEN
       #Control_Active := TRUE;

       #Temp_Error := #Temperature_SP - #Temperature_PV;

       #Control_Timer(IN := TRUE,
                      PT := #Control_Cycle);

       IF #Control_Timer.Q THEN
           //#Control_Timer(IN := FALSE,
                          //PT := T#0S);
           IF #Temp_Error > #Control_Deadband THEN
               // Need heating
               "DB_Valves".Valves[6].Open_Auto := TRUE;     // V6 steam
               "DB_Valves".Valves[9].Open_Auto := FALSE;    // V9 cooling
               "DB_Process".IO.DO_Steam_Regulator_En := TRUE;
               #Heating_Active := TRUE;

           ELSIF #Temp_Error < - #Control_Deadband THEN
               // Need cooling
               "DB_Valves".Valves[6].Open_Auto := FALSE;    // V6 steam
               "DB_Valves".Valves[9].Open_Auto := TRUE;     // V9 cooling
               "DB_Process".IO.DO_Cooling_Water := TRUE;
               #Cooling_Active := TRUE;

           ELSE
               // At setpoint
               "DB_Valves".Valves[6].Open_Auto := FALSE;
               "DB_Valves".Valves[9].Open_Auto := FALSE;
               "DB_Process".IO.DO_Steam_Regulator_En := FALSE;
               "DB_Process".IO.DO_Cooling_Water := FALSE;
           END_IF;
       END_IF;

       #At_Setpoint := ABS(#Temp_Error) <= #Control_Deadband;

       IF #At_Setpoint THEN
           #Status_Text := 'At setpoint';
       ELSIF #Heating_Active THEN
           #Status_Text := 'Heating active';
       ELSIF #Cooling_Active THEN
           #Status_Text := 'Cooling active';
       ELSE
           #Status_Text := 'Control active';
       END_IF;

   ELSE
       #Control_Active := FALSE;
       "DB_Valves".Valves[6].Open_Auto := FALSE;
       "DB_Valves".Valves[9].Open_Auto := FALSE;
       "DB_Process".IO.DO_Steam_Regulator_En := FALSE;
       "DB_Process".IO.DO_Cooling_Water := FALSE;
       #At_Setpoint := FALSE;
       #Control_Timer(IN := FALSE,
                      PT := T#0S);
       #Status_Text := 'Control disabled';
   END_IF;
END_FUNCTION_BLOCK

FUNCTION_BLOCK "FB_Vacuum_Controller"   // FB7, SCL
{ S7_Optimized_Access := 'TRUE' }
VERSION : 0.1
   VAR_INPUT
      Enable_Vacuum : Bool;
      Vacuum_Setpoint : Real;
      Pressure_PV : Real;
      Vacuum_Tolerance : Real;
      Safety_Permissive : Bool;
   END_VAR
   VAR_OUTPUT
      Vacuum_Active : Bool;
      At_Vacuum : Bool;
      Pump_Running : Bool;
      Status_Text : String;
   END_VAR
   VAR
      Pump_Start_Timer : TON_TIME;
      Pump_Stop_Timer : TON_TIME;
      Vacuum_Monitor : TON_TIME;
      Pump_Command : Bool;
      Vacuum_High_Limit : Real;
      Vacuum_Low_Limit : Real;
      Atmospheric_Press : Real := 1013.0;
   END_VAR
BEGIN
   #Vacuum_High_Limit := (#Atmospheric_Press - #Vacuum_Setpoint) + #Vacuum_Tolerance;
   #Vacuum_Low_Limit := (#Atmospheric_Press - #Vacuum_Setpoint) - #Vacuum_Tolerance;

   IF #Enable_Vacuum AND #Safety_Permissive THEN
       IF #Pressure_PV > #Vacuum_High_Limit THEN
           "DB_Valves".Valves[8].Open_Auto := TRUE;        // V8 vacuum
           "DB_Process".IO.DO_Vacuum_Pump := TRUE;
           #Pump_Start_Timer(IN := TRUE,
                             PT := T#5S);

           IF #Pump_Start_Timer.Q THEN
               #Pump_Running := TRUE;
               #Pump_Start_Timer(IN := FALSE,
                                 PT := T#0S);
           END_IF;
       ELSE
           "DB_Valves".Valves[8].Open_Auto := FALSE;
           "DB_Process".IO.DO_Vacuum_Pump := FALSE;
           #Pump_Running := FALSE;
       END_IF;

       #Vacuum_Active := "DB_Valves".Valves[8].Open_Auto;
       #At_Vacuum := (#Pressure_PV >= #Vacuum_Low_Limit) AND (#Pressure_PV <= #Vacuum_High_Limit);

       IF #At_Vacuum THEN
           #Status_Text := 'At vacuum setpoint';
       ELSIF #Vacuum_Active THEN
           #Status_Text := 'Pulling vacuum';
       ELSE
           #Status_Text := 'Vacuum ready';
       END_IF;

   ELSE
       #Vacuum_Active := FALSE;
       #Pump_Running := FALSE;
       #At_Vacuum := FALSE;
       "DB_Valves".Valves[8].Open_Auto := FALSE;
       "DB_Process".IO.DO_Vacuum_Pump := FALSE;
       #Status_Text := 'Vacuum system disabled';
   END_IF;
END_FUNCTION_BLOCK

FUNCTION_BLOCK "FB_Mixing_Phase"   // FB8, SCL
{ S7_Optimized_Access := 'TRUE' }
VERSION : 0.1
   VAR_INPUT
      Phase_Enable : Bool;
      Safety_Permissive : Bool;
      Reset_Phase : Bool;
   END_VAR
   VAR_OUTPUT
      Phase_Complete : Bool;
      Phase_Active : Bool;
      Phase_Fault : Bool;
      Phase_Status : String;
      Mixing_Active : Bool;
      Time_Remaining : Time;
      Phase_Progress : Real;
      Step_Status : String;
   END_VAR
   VAR_IN_OUT
      Motor_Controller : "FB_Motor_Controller";
   END_VAR
   VAR
      Mix_Timer : TON_TIME;
      Motor_FB_Instance : "FB_Motor_VFD";
   END_VAR
BEGIN
   IF #Reset_Phase THEN
       #Phase_Complete := FALSE;
       #Phase_Active := FALSE;
       #Phase_Fault := FALSE;
       #Phase_Status := 'Mixing phase reset';
       #Mixing_Active := FALSE;
       #Phase_Progress := 0.0;
       #Mix_Timer(IN := FALSE,
                  PT := T#0S);
       RETURN;
   END_IF;



   IF #Phase_Enable AND #Safety_Permissive AND "DB_Process".IO.Manhole_Closed_FB  THEN
       #Phase_Active := TRUE;
       #Phase_Status := 'Cold mixing active';
       #Mixing_Active := TRUE;
       #Step_Status:='Keep Manhole Closed';
       #Motor_Controller(
                         Enable := TRUE,
                         Command_Start := TRUE,

                         Speed_Setpoint := "DB_Recipes".Active_Recipe.Screw.Cold_Mix_Speed_pct,
                         Pulse_Enable := "DB_Recipes".Active_Recipe.Screw.Pulse_Enable_ColdMix,
                         Discharge_Mode := FALSE,
                         Direction_Command := 1,
                         Safety_Permissive := #Safety_Permissive,

                         Motor_FB := #Motor_FB_Instance
       );

       "DB_Valves".Valves[7].Open_Auto := TRUE;        // V7 evacuation
       "DB_Valves".Valves[2].Open_Auto := TRUE;
       "DB_Valves".Valves[3].Open_Auto := TRUE;

       #Mix_Timer(IN := TRUE,
                  PT := "DB_Recipes".Active_Recipe.Production.Cold_Mix_Time);
       #Time_Remaining := "DB_Recipes".Active_Recipe.Production.Cold_Mix_Time - #Mix_Timer.ET;

       IF "DB_Recipes".Active_Recipe.Production.Cold_Mix_Time > T#0S THEN
           #Phase_Progress := (DINT_TO_REAL(TIME_TO_DINT(#Mix_Timer.ET)) / DINT_TO_REAL(TIME_TO_DINT("DB_Recipes".Active_Recipe.Production.Cold_Mix_Time))) * 100.0;
       END_IF;

       IF #Mix_Timer.Q THEN
           #Phase_Complete := TRUE;
           #Phase_Active := FALSE;
           #Mixing_Active := FALSE;
           #Phase_Status := 'Cold mixing complete';

           #Motor_Controller.Command_Start := FALSE;
           "DB_Valves".Valves[7].Open_Auto := FALSE;
           "DB_Valves".Valves[3].Open_Auto := FALSE;
           "DB_Valves".Valves[2].Open_Auto := FALSE;
       END_IF;

   ELSE
       #Phase_Active := FALSE;
       #Phase_Complete := FALSE;
       #Mixing_Active := FALSE;
       #Mix_Timer(IN := FALSE,
                  PT := T#0S);

       #Motor_Controller.Command_Start := FALSE;
       "DB_Valves".Valves[7].Open_Auto := FALSE;
       "DB_Valves".Valves[3].Open_Auto := FALSE;
       "DB_Valves".Valves[2].Open_Auto := FALSE;
       #Phase_Status := 'Phase disabled';
   END_IF;
END_FUNCTION_BLOCK

FUNCTION_BLOCK "FB_Cooking_Phase"   // FB9, SCL
{ S7_Optimized_Access := 'TRUE' }
VERSION : 0.1
   VAR_INPUT
      Phase_Enable : Bool;
      Safety_Permissive : Bool;
      Reset_Phase : Bool;
   END_VAR
   VAR_OUTPUT
      Phase_Complete : Bool;
      Phase_Active : Bool;
      Phase_Fault : Bool;
      Step_Complete : Bool;
      Next_Step : UInt;
      Phase_Status : String;
      Step_Status : String;
      At_Temperature : Bool;
      Time_Remaining : Time;
      Phase_Progress : Real;
   END_VAR
   VAR_IN_OUT
      Motor_Controller : "FB_Motor_Controller";
      Temp_Controller : "FB_Temperature_Controller";
      Vacuum_Controller : "FB_Vacuum_Controller";
      Current_Step : UInt;
   END_VAR
   VAR
      Heating_Timer : TON_TIME;
      Cooking_Timer : TON_TIME;
      Motor_FB_Instance : "FB_Motor_VFD";
      Completed_Steps : UInt;
   END_VAR
BEGIN
   IF #Reset_Phase THEN
       #Phase_Complete := FALSE;
       #Phase_Active := FALSE;
       #Phase_Fault := FALSE;
       #Step_Complete := FALSE;
       #Phase_Status := 'Cooking phase reset';
       #Next_Step := 6;
       #Current_Step := #Next_Step;
       #Completed_Steps := 0;
       #Heating_Timer(IN := FALSE,
                      PT := T#0S);
       #Cooking_Timer(IN := FALSE,
                      PT := T#0S);
       "DB_Valves".Valves[2].Open_Auto := FALSE;
       "DB_Valves".Valves[3].Open_Auto := FALSE;
       "DB_Valves".Valves[6].Open_Auto := FALSE;
       "DB_Valves".Valves[9].Open_Auto := FALSE;
       "DB_Valves".Valves[8].Open_Auto := FALSE;
       RETURN;
   END_IF;

   IF #Phase_Enable AND #Safety_Permissive THEN
       #Phase_Active := TRUE;

       CASE #Current_Step OF
           6: // Heating Phase
               #Step_Status := 'Heating to setpoint';

               // Continue screw mixing
               #Motor_Controller(
                                 Enable := TRUE,
                                 Command_Start := TRUE,
                                 Speed_Setpoint := "DB_Recipes".Active_Recipe.Screw.Cook_Mix_Speed_pct,
                                 Pulse_Enable := "DB_Recipes".Active_Recipe.Screw.Pulse_Enable_Cooking,
                                 Discharge_Mode := FALSE,
                                 Direction_Command := 1,
                                 Safety_Permissive := #Safety_Permissive,

                                 Motor_FB := #Motor_FB_Instance
               );

               // Temperature control
               #Temp_Controller(
                                Enable_Control := TRUE,
                                Temperature_SP := "DB_Recipes".Active_Recipe.Temperature.Heat_Setpoint_Phase1,
                                Temperature_PV := "DB_Process".IO.AI_Temperature,
                                Control_Deadband := "DB_Recipes".Active_Recipe.Temperature.Heat_Deadband,
                                Safety_Permissive := #Safety_Permissive
               );

               #At_Temperature := #Temp_Controller.At_Setpoint;
               "DB_Valves".Valves[2].Open_Auto := TRUE;
               "DB_Valves".Valves[3].Open_Auto := TRUE;
               "DB_Valves".Valves[6].Open_Auto := TRUE;
               "DB_Valves".Valves[9].Open_Auto := TRUE;
               "DB_Valves".Valves[8].Open_Auto := TRUE;
               IF #At_Temperature THEN
                   #Step_Complete := TRUE;
                   #Next_Step := 7;
                   #Current_Step := #Next_Step;
                   #Completed_Steps := 1;
                   #Step_Status := 'Target temperature reached';
               END_IF;

           7: // Cooking Phase
               #Step_Status := 'Cooking at temperature';

               // Continue temperature and motor control
               #Temp_Controller(
                                Enable_Control := TRUE,
                                Temperature_SP := "DB_Recipes".Active_Recipe.Temperature.Heat_Setpoint_Phase1,
                                Temperature_PV := "DB_Process".IO.AI_Temperature,
                                Control_Deadband := "DB_Recipes".Active_Recipe.Temperature.Heat_Deadband,
                                Safety_Permissive := #Safety_Permissive
               );

               #Motor_Controller(
                                 Enable := TRUE,
                                 Command_Start := TRUE,
                                 Speed_Setpoint := "DB_Recipes".Active_Recipe.Screw.Cook_Mix_Speed_pct,
                                 Pulse_Enable := "DB_Recipes".Active_Recipe.Screw.Pulse_Enable_Cooking,
                                 Safety_Permissive := #Safety_Permissive,
                                 Motor_FB := #Motor_FB_Instance
               );

               // Vacuum if enabled
               IF "DB_Recipes".Active_Recipe.Vacuum.Cooking_Vacuum_Enable THEN
                   #Vacuum_Controller(
                                      Enable_Vacuum := TRUE,
                                      Vacuum_Setpoint := "DB_Recipes".Active_Recipe.Vacuum.Vacuum_Setpoint_mbar,
                                      Pressure_PV := "DB_Process".IO.AI_Pressure,
                                      Vacuum_Tolerance := "DB_Recipes".Active_Recipe.Vacuum.Vacuum_Tolerance,
                                      Safety_Permissive := #Safety_Permissive

                   );
               END_IF;

               // Cooking timer
               #Cooking_Timer(IN := TRUE,
                              PT := "DB_Recipes".Active_Recipe.Production.Cooking_Time_Phase1);
               #Time_Remaining := "DB_Recipes".Active_Recipe.Production.Cooking_Time_Phase1 - #Cooking_Timer.ET;

               IF "DB_Recipes".Active_Recipe.Production.Cooking_Time_Phase1 > T#0S THEN
                   #Phase_Progress := (DINT_TO_REAL(TIME_TO_DINT(#Cooking_Timer.ET)) / DINT_TO_REAL(TIME_TO_DINT("DB_Recipes".Active_Recipe.Production.Cooking_Time_Phase1))) * 100.0;
               END_IF;

               IF #Cooking_Timer.Q THEN
                   #Phase_Complete := TRUE;
                   #Step_Complete := TRUE;
                   #Next_Step := 10;  // Move to discharge phase
                   #Current_Step := #Next_Step;
                   "DB_Valves".Valves[2].Open_Auto := FALSE;
                   "DB_Valves".Valves[3].Open_Auto := FALSE;
                   "DB_Valves".Valves[6].Open_Auto := FALSE;
                   "DB_Valves".Valves[9].Open_Auto := FALSE;
                   "DB_Valves".Valves[8].Open_Auto := FALSE;
                   #Completed_Steps := 2;
                   #Phase_Status := 'Cooking complete';

               END_IF;

           ELSE
               #Phase_Fault := TRUE;
               #Phase_Status := 'Invalid cooking step';
       END_CASE;

   ELSE
       #Phase_Active := FALSE;
       #Phase_Complete := FALSE;
       #Phase_Status := 'Phase disabled';
   END_IF;
END_FUNCTION_BLOCK

FUNCTION_BLOCK "FB_Discharge_Phase"   // FB10, SCL
{ S7_Optimized_Access := 'TRUE' }
VERSION : 0.1
   VAR_INPUT
      Phase_Enable : Bool;
      Safety_Permissive : Bool;
      Reset_Phase : Bool;
   END_VAR
   VAR_OUTPUT
      Phase_Complete : Bool;
      Phase_Active : Bool;
      Phase_Fault : Bool;
      Step_Complete : Bool;
      Next_Step : UInt;
      Phase_Status : String;
      Step_Status : String;
      Discharge_Active : Bool;
      Ready_For_Discharge : Bool;
      Time_Remaining : Time;
      Phase_Progress : Real;
   END_VAR
   VAR_IN_OUT
      Motor_Controller : "FB_Motor_Controller";
      Current_Step : UInt;
   END_VAR
   VAR
      Discharge_Timer : TON_TIME;
      Confirm_Timer : TON_TIME;
      Discharge_Started : Bool;
      Total_Steps : UInt := 3;
      Completed_Steps : UInt;
      Motor_FB_Instance : "FB_Motor_VFD";
   END_VAR
BEGIN
   #Phase_Complete := FALSE;

   IF #Reset_Phase THEN
       #Phase_Complete := FALSE;
       #Phase_Active := FALSE;
       #Phase_Fault := FALSE;
       #Step_Complete := FALSE;
       #Phase_Status := 'Discharge phase reset';
       #Discharge_Active := FALSE;
       #Ready_For_Discharge := FALSE;
       #Next_Step := 10;
       #Current_Step := #Next_Step;
       #Completed_Steps := 0;
       #Discharge_Timer(IN := FALSE,
                        PT := T#0S);
       #Confirm_Timer(IN := FALSE,
                      PT := T#0S);
       RETURN;
   END_IF;

   IF #Phase_Enable AND #Safety_Permissive THEN
       #Phase_Active := TRUE;

       CASE #Current_Step OF
           10: // Wait to Confirm Discharge
               #Phase_Status := 'Discharging phase';
               #Step_Status := 'Awaiting discharge confirm';

               #Ready_For_Discharge := TRUE;

               "DB_Valves".Valves[6].Open_Auto := FALSE;       // V6 Steam OFF
               "DB_Valves".Valves[2].Open_Auto := TRUE;        // V4 Discharge
               "DB_Valves".Valves[3].Open_Auto := TRUE;
               #Motor_Controller(
                                 Enable := TRUE,
                                 Command_Start := TRUE,
                                 Speed_Setpoint := 30.0,
                                 Pulse_Enable := FALSE,
                                 Discharge_Mode := FALSE,
                                 Direction_Command := 1,
                                 Safety_Permissive := #Safety_Permissive,

                                 Motor_FB := #Motor_FB_Instance
               );

               #Confirm_Timer(IN := TRUE,
                              PT := T#30S);

               IF "DB_Process".HMI.Discharge_Ready_OK THEN
                   #Step_Complete := TRUE;
                   #Next_Step := 11;
                   #Current_Step := #Next_Step;
                   #Completed_Steps := 1;
                   #Ready_For_Discharge := FALSE;
               ELSIF #Confirm_Timer.Q THEN
                   #Phase_Fault := TRUE;
                   #Step_Status := 'Discharge confirm timeout';
               END_IF;

           11: // Discharge Product
               #Step_Status := 'Discharging product';
               #Discharge_Active := TRUE;

               "DB_Valves".Valves[2].Open_Auto := TRUE;        // V4 Discharge
               "DB_Valves".Valves[4].Open_Auto := TRUE;        // V3 Unlock

               #Motor_Controller(
                                 Enable := TRUE,
                                 Command_Start := TRUE,
                                 Speed_Setpoint := "DB_Recipes".Active_Recipe.Screw.Discharge_Speed_pct,
                                 Pulse_Enable := "DB_Recipes".Active_Recipe.Screw.Pulse_Enable_Discharge,
                                 Discharge_Mode := TRUE,
                                 Direction_Command := 1,
                                 Safety_Permissive := #Safety_Permissive,

                                 Motor_FB := #Motor_FB_Instance
               );

               IF "DB_Recipes".Active_Recipe.Production.Discharge_Time > T#0S THEN
                   #Discharge_Timer(IN := TRUE,
                                    PT := "DB_Recipes".Active_Recipe.Production.Discharge_Time);
                   #Time_Remaining := "DB_Recipes".Active_Recipe.Production.Discharge_Time - #Discharge_Timer.ET;

                   IF #Discharge_Timer.Q THEN
                       #Step_Complete := TRUE;
                       #Next_Step := 12;
                       #Current_Step := #Next_Step;

                       #Completed_Steps := 2;
                   END_IF;

                   #Phase_Progress := (DINT_TO_REAL(TIME_TO_DINT(#Discharge_Timer.ET)) / DINT_TO_REAL(TIME_TO_DINT("DB_Recipes".Active_Recipe.Production.Discharge_Time))) * 100.0;
               ELSE
                   #Step_Status := 'Manual discharge active';
                   #Discharge_Timer(IN := TRUE,
                                    PT := T#6S);
                   IF #Discharge_Timer.Q THEN
                       #Step_Complete := TRUE;
                       #Next_Step := 12;
                       #Current_Step := #Next_Step;
                       #Completed_Steps := 2;
                   END_IF;
               END_IF;

           12: // Finalize
               #Step_Status := 'Finalizing batch';
               #Discharge_Active := FALSE;

               #Motor_Controller(
                                 Enable := FALSE,
                                 Command_Start := FALSE,
                                 Speed_Setpoint := 0.0,
                                 Pulse_Enable := FALSE,
                                 Discharge_Mode := FALSE,
                                 Direction_Command := 0,
                                 Safety_Permissive := FALSE,

                                 Motor_FB := #Motor_FB_Instance
               );

               // Turn off all valves
               "DB_Valves".Valves[4].Open_Auto := FALSE;       // V4 Discharge
               "DB_Valves".Valves[6].Open_Auto := FALSE;       // V6 Steam
               "DB_Valves".Valves[7].Open_Auto := FALSE;       // V7 Evacuation
               "DB_Valves".Valves[8].Open_Auto := FALSE;       // V8 Vacuum
               "DB_Valves".Valves[3].Open_Auto := FALSE;       // V3 Unlock
               "DB_Valves".Valves[3].Close_Auto := FALSE;       // V3 Unlock
               "DB_Valves".Valves[2].Open_Auto := FALSE;       // V3 Unlock

               #Phase_Complete := TRUE;
               #Phase_Active := FALSE;
               #Completed_Steps := 3;
               #Phase_Status := 'Batch complete';
               #Phase_Progress := 100.0;




           ELSE
               #Phase_Fault := TRUE;
               #Phase_Status := 'Invalid discharge step';
       END_CASE;

       IF NOT #Phase_Complete THEN
           #Phase_Progress := (UINT_TO_REAL(#Completed_Steps) / UINT_TO_REAL(#Total_Steps)) * 100.0;
       END_IF;

   ELSE
       #Phase_Active := FALSE;
       #Phase_Complete := FALSE;
       #Phase_Status := 'Phase disabled';
   END_IF;
END_FUNCTION_BLOCK

FUNCTION_BLOCK "FB_Process_Main"   // FB11, SCL
{ S7_Optimized_Access := 'TRUE' }
VERSION : 0.1
   VAR_OUTPUT
      Process_Running : Bool;
      Current_Step : UInt;
      Current_Phase : UInt;
      System_Ready : Bool;
      Status_Message : String;
      Phase_Message : String;
      phase_Progress : Real;
      Fault_Text : String;
      Fault_Code : UInt;
   END_VAR
   VAR
      Motor_Controller : "FB_Motor_Controller";
      Motor_FB_Instance : "FB_Motor_VFD";
      Temp_Controller : "FB_Temperature_Controller";
      Vacuum_Controller : "FB_Vacuum_Controller";
      Preparation_Phase : "FB_Preparation_Phase";
      Mixing_Phase : "FB_Mixing_Phase";
      Cooking_Phase : "FB_Cooking_Phase";
      Discharge_Phase : "FB_Discharge_Phase";
      Internal_Step : UInt;
      Safety_OK : Bool;
      Recipe_Loaded : Bool;
      Prep_Complete : Bool;
      Mix_Complete : Bool;
      Cook_Complete : Bool;
      Discharge_Complete : Bool;
      First_Scan : Bool := True;
      Individual_Discharge_Active : Bool;
      Individual_Discharge_Timer : TON_TIME;
      Individual_Discharge_Enable : Bool;
   END_VAR
   VAR_TEMP
      Temp_Emergency_Active : Bool;
   END_VAR
BEGIN
   // Initialize outputs
   #Process_Running := FALSE;
   #System_Ready := FALSE;
   #Status_Message := '';
   #Phase_Message := '';

   IF #First_Scan THEN
       "DB_Process".Status.Current_Step := 50;
       "DB_Process".Status.Current_Phase := 0;
       #First_Scan := FALSE;
   END_IF;




   // Read current state
   #Current_Step := "DB_Process".Status.Current_Step;
   #Current_Phase := "DB_Process".Status.Current_Phase;

   // Safety monitoring
   "FC_Safety_Monitor"(
                       Emergency_Stop := "DB_Process".IO.ES_Emergency_Stop,
                       Door_Interlock_OK := "DB_Process".IO.Door_Interlock_OK,
                       Door_Locked:="DB_Process".IO.Door_Locked_FB,
                       Manhole_Secured:="DB_Process".IO.Manhole_Closed_FB,
                       Temperature_Value := "DB_Process".IO.AI_Temperature,
                       Pressure_Value := "DB_Process".IO.AI_Pressure,
                       System_Enabled := TRUE,

                       Safety_OK => #Safety_OK,
                       System_Ready => #System_Ready,
                       Emergency_Active=>#Temp_Emergency_Active,
                       Safety_Fault => "DB_Process".Status.Fault_Active,
                       Fault_Code=>#Fault_Code,
                       Fault_Text=>#Fault_Text
   );

   // Process control
   IF "DB_Process".IO.ES_Emergency_Stop THEN
       #Current_Phase := 0;
       #Current_Step := 99;
       #Status_Message := 'EMERGENCY STOP ACTIVE';
       #Process_Running := FALSE;

   ELSIF "DB_Process".HMI.Reset_System THEN
       #Current_Phase := 0;
       #Current_Step := 50;
       #Status_Message := 'System reset';
       #Process_Running := FALSE;
       "DB_Process".HMI.Start_Production := FALSE;
       "DB_Process".IO.Water_Level_FB:=FALSE;
       "DB_Process".IO.Door_Locked_FB := FALSE;
       "DB_Process".IO.Door_Interlock_OK := FALSE;
       "DB_Process".IO.Manhole_Closed_FB := FALSE;
       "DB_Process".IO.Manhole_Open_FB := TRUE;
       #Prep_Complete := FALSE;
       #Mix_Complete := FALSE;
       #Cook_Complete := FALSE;
       #Discharge_Complete := FALSE;

   ELSIF "DB_Process".HMI.Start_Production AND #Safety_OK THEN
       #Process_Running := TRUE;
       IF #Current_Phase = 0 THEN
           #Current_Phase := 1;
           #Current_Step := 15;
           #Status_Message := 'Process started';
       END_IF;

   ELSIF "DB_Process".HMI.Stop_Production THEN
       #Process_Running := FALSE;
       #Status_Message := 'Process stopped';
   END_IF;

   // Main phase coordination with ALL controllers
   IF #Process_Running AND #Safety_OK THEN
       CASE #Current_Phase OF
           1: // Preparation Phase (Steps 15→1→2→3→4)
               #Preparation_Phase(
                                  Phase_Enable := TRUE,
                                  Current_Step := #Current_Step,
                                  Safety_Permissive := #Safety_OK,
                                  Reset_Phase := "DB_Process".HMI.Reset_p_s, // add reset phase button

                                  Phase_Complete => #Prep_Complete,
                                  Next_Step => #Internal_Step,
                                  Step_Status=> #Status_Message,
                                  Phase_Status => #Phase_Message,
                                  Phase_Progress=>#phase_Progress

               );


               IF #Prep_Complete THEN
                   #Current_Phase := 2;
                   #Current_Step := 5;
               END_IF;

           2: // Mixing Phase (Step 5)
               #Mixing_Phase(
                             Phase_Enable := TRUE,
                             Safety_Permissive := #Safety_OK,
                             Reset_Phase := "DB_Process".HMI.Reset_p_s,

                             Motor_Controller := #Motor_Controller,

                             Phase_Complete => #Mix_Complete,
                             Step_Status=> #Status_Message,
                               Phase_Status => #Phase_Message,
                             Phase_Progress=>#phase_Progress
               );


               IF #Mix_Complete THEN
                   #Current_Phase := 3;
                   #Current_Step := 6;
               END_IF;

           3: // Cooking Phase (Steps 6→7)
               #Cooking_Phase(
                              Phase_Enable := TRUE,
                              Current_Step := #Current_Step,
                              Safety_Permissive := #Safety_OK,
                              Reset_Phase := "DB_Process".HMI.Reset_p_s,

                              Motor_Controller := #Motor_Controller,
                              Temp_Controller := #Temp_Controller,
                              Vacuum_Controller := #Vacuum_Controller,

                              Phase_Complete => #Cook_Complete,
                              Next_Step => #Internal_Step,

                              Phase_Status => #Phase_Message,
                              Step_Status=>#Status_Message,
                              Phase_Progress =>#phase_Progress
               );

               #Current_Step := #Internal_Step;

               IF #Cook_Complete THEN
                   #Current_Phase := 4;
                   #Current_Step := 10;
               END_IF;

           4: // Discharge Phase (Steps 10→11→12)
               #Discharge_Phase(
                                Phase_Enable := TRUE,
                                Current_Step := #Current_Step,
                                Safety_Permissive := #Safety_OK,
                                Reset_Phase := "DB_Process".HMI.Reset_p_s,

                                Motor_Controller := #Motor_Controller,

                                Phase_Complete => #Discharge_Complete,
                                Next_Step => #Internal_Step,
                                Phase_Status => #Phase_Message,
                                Step_Status=>#Status_Message,
                                Phase_Progress =>#phase_Progress
               );
               #Current_Step := #Internal_Step;

               IF #Discharge_Complete THEN
                   #Process_Running := FALSE;
                   #Current_Phase := 0;
                   #Current_Step := 50;
                   "DB_Process".IO.Door_Locked_FB := FALSE;
                   "DB_Process".IO.Manhole_Closed_FB := false;
                   "DB_Process".IO.Manhole_Open_FB := TRUE;
                   "DB_Process".IO.Water_Level_FB := False;
                   "DB_Process".IO.Door_Interlock_OK := False;
                   "DB_Process".HMI.Individual_Discharge_Button := False;


                   #Status_Message := 'PROCESS COMPLETE - BATCH FINISHED';
               END_IF;

           ELSE
               #Status_Message := 'Invalid phase';
       END_CASE;

   ELSE
       #Status_Message := 'System idle - ready for operation';
   END_IF;

   // ===== INDIVIDUAL DISCHARGE BUTTON LOGIC =====
   // Individual discharge can only run when process is NOT running
   IF "DB_Process".HMI.Individual_Discharge_Button AND
       NOT "DB_Process".Status.Process_Running AND
       #Safety_OK THEN
       #Individual_Discharge_Active := TRUE;
       #Individual_Discharge_Enable := TRUE;
       // Start discharge sequence
       "DB_Valves".Valves[4].Open_Auto := TRUE; // V4 Discharge valve
       "DB_Valves".Valves[3].Open_Auto := TRUE; // V3 Unlock valve
       // Start motor at discharge speed
       "DB_Motors".Motors[1].Command.Start_Auto := TRUE;
       "DB_Motors".Motors[1].Command.Speed_SP_pct := 25.0;
       "DB_Motors".Motors[1].Command.Discharge_Mode := TRUE;
       // Safety timer - maximum 10 minutes
       #Individual_Discharge_Timer(IN := TRUE,
                                   PT := T#600S);
       // Stop if timer expires
       IF #Individual_Discharge_Timer.Q THEN
           #Individual_Discharge_Active := FALSE;
       END_IF;
   ELSE
       #Individual_Discharge_Active := FALSE;
       #Individual_Discharge_Enable := FALSE;
       #Individual_Discharge_Timer(IN := FALSE,
                                   PT := T#0S);
       // Stop individual discharge only if process is not running
       IF NOT "DB_Process".Status.Process_Running THEN
           "DB_Valves".Valves[4].Open_Auto := FALSE;
           "DB_Valves".Valves[3].Open_Auto := FALSE;
           "DB_Motors".Motors[1].Command.Start_Auto := FALSE;
           "DB_Motors".Motors[1].Command.Discharge_Mode := FALSE;
       END_IF;
   END_IF;
   // Update status
   "DB_Process".Status.Individual_Discharge_Active := #Individual_Discharge_Active;

   // Update process status
   "DB_Process".Status.Current_Step := #Current_Step;
   "DB_Process".Status.Current_Phase := #Current_Phase;
   "DB_Process".Status.Process_Running := #Process_Running;
   "DB_Process".Status.System_Ready := #System_Ready;
   "DB_Process".Status.Step_Name := #Status_Message;
   "DB_Process".Status.Phase_Name := #Phase_Message;
END_FUNCTION_BLOCK

FUNCTION_BLOCK "FB_Valve_Controller"   // FB12, SCL
{ S7_Optimized_Access := 'TRUE' }
VERSION : 0.1
   VAR_INPUT
      Open_Command : Bool;
      Enable : Bool;
      Close_Command : Bool;
      Safety_Permissive : Bool;
      Emergency_Close : Bool;
      Position_SP : Real;
   END_VAR
   VAR_OUTPUT
      Valve_Open : Bool;
      Valve_Closed : Bool;
      Valve_Ready : Bool;
      Valve_Fault : Bool;
      Status_Text : String;
   END_VAR
   VAR_IN_OUT
      Valve_Data : "UDT_Valve";
      Valve_FB : "FB_Valve_DO";
   END_VAR
   VAR
      Temp_Position : Real;
      Temp_Operation_Count : UDInt;
      Temp_Runtime : Real;
   END_VAR
BEGIN
   // Set commands based on inputs
   IF #Enable AND #Safety_Permissive THEN
       #Valve_Data.Open_Auto := #Open_Command
       ;
       #Valve_Data.Close_Auto := #Close_Command
       ;
       #Valve_Data.Enable := TRUE;
   ELSE
       #Valve_Data.Open_Auto := FALSE;
       #Valve_Data.Close_Auto := FALSE;
       #Valve_Data.Enable := FALSE;
   END_IF;

   // Set interlocks
   #Valve_Data.Interlocks.Permissive := #Safety_Permissive;
   #Valve_Data.Interlocks.OOS := NOT #Enable;
   #Valve_Data.Interlocks.E_Stop := "DB_Process".IO.ES_Emergency_Stop;

   // Call valve FB
   #Valve_FB(
             ManCmd := #Valve_Data.Open_Man,
             FuncCmd := #Valve_Data.Open_Func,
             AutoCmd := #Valve_Data.Open_Auto,

             Permissive := #Valve_Data.Interlocks.Permissive,
             OOS := #Valve_Data.Interlocks.OOS,

             Q_Open => #Valve_Data.Outputs.Q_Open,
             Q_Close => #Valve_Data.Outputs.Q_Close,
             Ready => #Valve_Data.Status.Ready

             // Assign unused outputs to temp variables

   );

   // Set outputs
   #Valve_Open := #Valve_Data.Status.Open;
   #Valve_Closed := #Valve_Data.Status.Closed;
   #Valve_Ready := #Valve_Data.Status.Ready;
   #Valve_Fault := #Valve_Data.Status.Fault;

   IF #Valve_Fault THEN
       #Status_Text := 'Valve fault';
   ELSIF #Valve_Open THEN
       #Status_Text := 'Open';
   ELSIF #Valve_Closed THEN
       #Status_Text := 'Closed';
   ELSE
       #Status_Text := 'Moving';
   END_IF;
END_FUNCTION_BLOCK

FUNCTION "FC_Test_Setup" : Void   // FC1, LAD
{ S7_Optimized_Access := 'FALSE' }
VERSION : 0.1
BEGIN

REGION Network 1
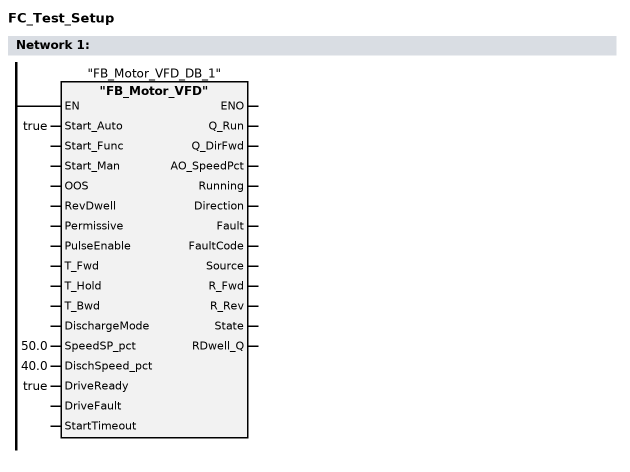
   RUNG wire#powerrail
      "FB_Motor_VFD_DB_1"(Start_Auto := true, Start_Func :=, Start_Man :=, OOS :=, RevDwell :=, Permissive :=, PulseEnable :=, T_Fwd :=, T_Hold :=, T_Bwd :=, DischargeMode :=, SpeedSP_pct := 50.0, DischSpeed_pct := 40.0, DriveReady := true, DriveFault :=, StartTimeout :=, Q_Run =>, Q_DirFwd =>, AO_SpeedPct =>, Running =>, Direction =>, Fault =>, FaultCode =>, Source =>, R_Fwd =>, R_Rev =>, State =>, RDwell_Q =>)
   END_RUNG
   // the same network as SCL:
   "FB_Motor_VFD_DB_1"(Start_Auto := true, SpeedSP_pct := 50.0, DischSpeed_pct := 40.0, DriveReady := true);   // "FB_Motor_VFD"
END_REGION
END_FUNCTION

FUNCTION "FC_Analog_Scaling" : Void   // FC2, SCL
{ S7_Optimized_Access := 'TRUE' }
VERSION : 0.1
   VAR_INPUT
      Raw_Value : Word;   // // Raw analog input (0-27648)
      Min_EU : Real;   // // Minimum engineering unit
      Max_EU : Real;   // // Maximum engineering unit
      Raw_Min : Word;   // // Raw minimum value (default 0)
      Raw_Max : Word;   // Raw maximum value (default 27648)
   END_VAR
   VAR_OUTPUT
      Scaled_Value : Real;   // / Scaled engineering value
      Valid : Bool;   // Value is within valid range
      Out_of_Range : Bool;
   END_VAR
   VAR_TEMP
      Raw_Value_DINT : DInt;
      Raw_Min_DINT : DInt;
      Raw_Max_DINT : DInt;
      Raw_Span_REAL : Real;
      Raw_Offset_REAL : Real;
      EU_Span : Real;
   END_VAR
BEGIN
   // Input validation
   IF #Raw_Value < #Raw_Min OR #Raw_Value > #Raw_Max THEN
       #Valid := FALSE;
       #Out_of_Range := TRUE;
       #Scaled_Value := 0.0;
       RETURN;
   END_IF;

   // Convert to DINT to avoid overflow (CORRECTED)
   #Raw_Value_DINT := WORD_TO_DINT(#Raw_Value);
   #Raw_Min_DINT := WORD_TO_DINT(#Raw_Min);
   #Raw_Max_DINT := WORD_TO_DINT(#Raw_Max);

   // Convert to REAL for calculations
   #Raw_Offset_REAL := DINT_TO_REAL(#Raw_Value_DINT - #Raw_Min_DINT);
   #Raw_Span_REAL := DINT_TO_REAL(#Raw_Max_DINT - #Raw_Min_DINT);
   #EU_Span := #Max_EU - #Min_EU;

   // Scaling calculation
   IF #Raw_Span_REAL > 0.0 THEN
       #Scaled_Value := #Min_EU + ((#Raw_Offset_REAL / #Raw_Span_REAL) * #EU_Span);
       #Valid := TRUE;
       #Out_of_Range := FALSE;
   ELSE
       #Valid := FALSE;
       #Out_of_Range := FALSE;
       #Scaled_Value := #Min_EU;
   END_IF;
END_FUNCTION

FUNCTION "FC_Motor_Integration" : Void   // FC3, SCL
{ S7_Optimized_Access := 'TRUE' }
VERSION : 0.1
   VAR_INPUT
      Motor_Number : UInt;
   END_VAR
   VAR_OUTPUT
      Integration_OK : Bool;
   END_VAR
   VAR_IN_OUT
      Motor_Data : "UDT_Motor";
      Motor_FB_Instance : "FB_Motor_VFD";
   END_VAR
BEGIN
   // Configure motor parameters for screw operation
   #Motor_Data.Config.Motor_Name := 'SCREW_MOTOR';
   #Motor_Data.Config.T_Fwd := #Motor_Data.Config.T_Fwd;        // From recipe
   #Motor_Data.Config.T_Hold := #Motor_Data.Config.T_Hold;      // From recipe  
   #Motor_Data.Config.T_Bwd := #Motor_Data.Config.T_Bwd;        // From recipe
   #Motor_Data.Config.Disch_Speed_pct := #Motor_Data.Config.Disch_Speed_pct;

   // Map UDT commands to your FB inputs
   #Motor_FB_Instance(
                      // Command inputs
                      Start_Man := #Motor_Data.Command.Start_Man,
                      Start_Func := #Motor_Data.Command.Start_Func,
                      Start_Auto := #Motor_Data.Command.Start_Auto,
                      OOS := #Motor_Data.Interlocks.OOS,
                      RevDwell := #Motor_Data.Config.Rev_Dwell,
                      Permissive := #Motor_Data.Interlocks.Permissive,
                      PulseEnable := #Motor_Data.Command.Pulse_Enable,
                      T_Fwd := #Motor_Data.Config.T_Fwd,
                      T_Hold := #Motor_Data.Config.T_Hold,
                      T_Bwd := #Motor_Data.Config.T_Bwd,
                      DischargeMode := #Motor_Data.Command.Discharge_Mode,
                      SpeedSP_pct := #Motor_Data.Command.Speed_SP_pct,
                      DischSpeed_pct := #Motor_Data.Config.Disch_Speed_pct,
                      DriveReady := #Motor_Data.Interlocks.Drive_Ready,
                      DriveFault := #Motor_Data.Interlocks.Drive_Fault,
                      StartTimeout := #Motor_Data.Config.Start_Timeout,

                      // Output mappings
                      Q_Run => #Motor_Data.Outputs.Q_Run,
                      Q_DirFwd => #Motor_Data.Outputs.Q_DirFwd,
                      AO_SpeedPct => #Motor_Data.Outputs.AO_SpeedPct,
                      Running => #Motor_Data.Status.Running,
                      Direction => #Motor_Data.Status.Direction,
                      Fault => #Motor_Data.Status.Fault,
                      FaultCode => #Motor_Data.Status.Fault_Code,
                      Source => #Motor_Data.Status.Source,
                      R_Fwd => #Motor_Data.Status.R_Fwd,
                      R_Rev => #Motor_Data.Status.R_Rev,
                      State => #Motor_Data.Status.State,
                      RDwell_Q => #Motor_Data.Status.RDwell_Q
   );

   // Set integration status
   #Integration_OK := TRUE;
END_FUNCTION

FUNCTION "FC_Timer_Manager" : Void   // FC4, SCL
{ S7_Optimized_Access := 'TRUE' }
VERSION : 0.1
   VAR_INPUT
      Timer_ID : UInt;   // // Timer ID (1-20)
      Start_Timer : Bool;
      Reset_Timer : Bool;
      Timer_PT : Time;   // // Timer preset time
   END_VAR
   VAR_OUTPUT
      Timer_Q : Bool;   // // Timer output (done)
      Timer_ET : Time;   // // Timer elapsed time
      Timer_Valid : Bool;   // // Timer ID is valid
   END_VAR
   VAR_IN_OUT
      Timer_Array : Array[1..20] of TON_TIME;
   END_VAR
BEGIN
   // Validate timer ID
   IF #Timer_ID < 1 OR #Timer_ID > 20 THEN
       #Timer_Valid := FALSE;
       #Timer_Q := FALSE;
       #Timer_ET := T#0S;
       RETURN;
   END_IF;

   #Timer_Valid := TRUE;

   // Timer control
   IF #Reset_Timer THEN
       #Timer_Array[#Timer_ID](IN := FALSE,
                               PT := T#0S);
   ELSE
       #Timer_Array[#Timer_ID](IN := #Start_Timer,
                               PT := #Timer_PT);
   END_IF;

   // Outputs
   #Timer_Q := #Timer_Array[#Timer_ID].Q;
   #Timer_ET := #Timer_Array[#Timer_ID].ET;
END_FUNCTION

FUNCTION "FC_Recipe_Manager" : Void   // FC5, SCL
{ S7_Optimized_Access := 'TRUE' }
VERSION : 0.1
   VAR_INPUT
      Recipe_Number : UInt;
      Load_Command : Bool;
      Save_Command : Bool;
      Validate_Command : Bool;
   END_VAR
   VAR_OUTPUT
      Operation_OK : Bool;
      Recipe_Valid : Bool;
      Error_Code : UInt;
      Error_Text : String;
   END_VAR
   VAR_IN_OUT
      Temp_Recipe : "UDT_Recipe_Complete";
   END_VAR
   VAR_TEMP
      RetVal : Int;
      Temp_DT : DTL;
      Status : Int;
   END_VAR
BEGIN
   // Initialize outputs
   #Operation_OK := FALSE;
   #Recipe_Valid := FALSE;
   #Error_Code := 0;
   #Error_Text := '';

   // Validate recipe number
   IF #Recipe_Number < 1 OR #Recipe_Number > 10 THEN
       #Error_Code := 101;
       #Error_Text := 'Invalid recipe number (1-10)';
       RETURN;
   END_IF;



   // Load recipe
   IF #Load_Command THEN
       #Temp_Recipe := "DB_Recipes".Recipes[#Recipe_Number];
       "DB_Recipes".Active_Recipe := #Temp_Recipe;
       #Operation_OK := TRUE;
       #Recipe_Valid := TRUE;
       #Error_Text := 'Recipe loaded successfully';
   END_IF;

   // Save recipe  
   IF #Save_Command THEN
       #Temp_Recipe := "DB_Recipes".Active_Recipe;
       #Status := RD_SYS_T(#Temp_DT);
       #Temp_Recipe.Modified_Date := #Temp_DT;

       #Temp_Recipe.Modified_By := 'OPERATOR';

       "DB_Recipes".Recipes[#Recipe_Number] := #Temp_Recipe;
       #Operation_OK := TRUE;
       #Error_Text := 'Recipe saved successfully';
   END_IF;

   // Validate recipe parameters
   IF #Validate_Command THEN
       #Temp_Recipe := "DB_Recipes".Active_Recipe;
       #Recipe_Valid := TRUE;

       // Check production parameters
       IF #Temp_Recipe.Production.Heating_Temp_Phase1 <= 0.0 OR
           #Temp_Recipe.Production.Heating_Temp_Phase1 > 100.0 THEN
           #Recipe_Valid := FALSE;
           #Error_Code := 201;
           #Error_Text := 'Invalid heating temperature (0-100C)';
       END_IF;

       // Check screw parameters
       IF #Temp_Recipe.Screw.Forward_Speed_pct < 0.0 OR
           #Temp_Recipe.Screw.Forward_Speed_pct > 100.0 THEN
           #Recipe_Valid := FALSE;
           #Error_Code := 202;
           #Error_Text := 'Invalid forward speed (0-100%)';
       END_IF;

       // Check times
       IF #Temp_Recipe.Production.Cold_Mix_Time <= T#0S THEN
           #Recipe_Valid := FALSE;
           #Error_Code := 203;
           #Error_Text := 'Invalid cold mix time';
       END_IF;

